screen "Lists" 1440x900, template "Tpl"
   TextField "frm_1" at 12,128 size 1416x70; Text 'Text'
   TextField "txt_1" at 21,132 size 300x23; Text 'POSTAVKE (dok sustav stoji)'
   TextField "txt_2" at 21,162 size 120x28; Text 'Redoslijed'
   SymbolicIOField "sym_1" at 141,162 size 248x28; TextOff '0'; TextOn '1'; TextList "TL_Order"
      ProcessValue <- "CfgOrderMode"
   TextField "txt_3" at 420,162 size 218x28; Text 'SEMI: transfer po koraku'
   SymbolicIOField "sym_2" at 638,162 size 82x28; TextOff '0'; TextOn '1'; TextList "TL_YesNo"
      ProcessValue <- "CfgSemiPerTransfer"
   TextField "txt_4" at 750,162 size 135x28; Text 'Ravnoteža'
   SymbolicIOField "sym_3" at 885,162 size 195x28; TextOff '0'; TextOn '1'; TextList "TL_BalMode"
      ProcessValue <- "CfgBalMode"
   TextField "txt_5" at 1110,162 size 60x28; Text 'Istovar'
   IOField "io_1" at 1170,162 size 45x28; FormatPattern 99
      ProcessValue <- "UTotal"
   TextField "txt_6" at 1230,162 size 60x28; Text 'Ukrcaj'
   IOField "io_2" at 1290,162 size 45x28; FormatPattern 99
      ProcessValue <- "LTotal"
   TextField "txt_7" at 12,210 size 350x23; Text 'LISTA ZA ISTOVAR (DB20) 1-24'
   TextField "txt_8" at 12,238 size 34x22; Text '1'
   IOField "io_3" at 51,238 size 68x22; FormatPattern 999
      ProcessValue <- "UList_01"
   SymbolicIOField "sym_4" at 123,238 size 112x22; TextOff '0'; TextOn '1'; TextList "TL_ListSt"
      ProcessValue <- "UState_01"
   TextField "txt_9" at 12,263 size 34x22; Text '2'
   IOField "io_4" at 51,263 size 68x22; FormatPattern 999
      ProcessValue <- "UList_02"
   SymbolicIOField "sym_5" at 123,263 size 112x22; TextOff '0'; TextOn '1'; TextList "TL_ListSt"
      ProcessValue <- "UState_02"
   TextField "txt_10" at 12,288 size 34x22; Text '3'
   IOField "io_5" at 51,288 size 68x22; FormatPattern 999
      ProcessValue <- "UList_03"
   SymbolicIOField "sym_6" at 123,288 size 112x22; TextOff '0'; TextOn '1'; TextList "TL_ListSt"
      ProcessValue <- "UState_03"
   TextField "txt_11" at 12,313 size 34x22; Text '4'
   IOField "io_6" at 51,313 size 68x22; FormatPattern 999
      ProcessValue <- "UList_04"
   SymbolicIOField "sym_7" at 123,313 size 112x22; TextOff '0'; TextOn '1'; TextList "TL_ListSt"
      ProcessValue <- "UState_04"
   TextField "txt_12" at 12,338 size 34x22; Text '5'
   IOField "io_7" at 51,338 size 68x22; FormatPattern 999
      ProcessValue <- "UList_05"
   SymbolicIOField "sym_8" at 123,338 size 112x22; TextOff '0'; TextOn '1'; TextList "TL_ListSt"
      ProcessValue <- "UState_05"
   TextField "txt_13" at 12,363 size 34x22; Text '6'
   IOField "io_8" at 51,363 size 68x22; FormatPattern 999
      ProcessValue <- "UList_06"
   SymbolicIOField "sym_9" at 123,363 size 112x22; TextOff '0'; TextOn '1'; TextList "TL_ListSt"
      ProcessValue <- "UState_06"
   TextField "txt_14" at 12,388 size 34x22; Text '7'
   IOField "io_9" at 51,388 size 68x22; FormatPattern 999
      ProcessValue <- "UList_07"
   SymbolicIOField "sym_10" at 123,388 size 112x22; TextOff '0'; TextOn '1'; TextList "TL_ListSt"
      ProcessValue <- "UState_07"
   TextField "txt_15" at 12,413 size 34x22; Text '8'
   IOField "io_10" at 51,413 size 68x22; FormatPattern 999
      ProcessValue <- "UList_08"
   SymbolicIOField "sym_11" at 123,413 size 112x22; TextOff '0'; TextOn '1'; TextList "TL_ListSt"
      ProcessValue <- "UState_08"
   TextField "txt_16" at 12,438 size 34x22; Text '9'
   IOField "io_11" at 51,438 size 68x22; FormatPattern 999
      ProcessValue <- "UList_09"
   SymbolicIOField "sym_12" at 123,438 size 112x22; TextOff '0'; TextOn '1'; TextList "TL_ListSt"
      ProcessValue <- "UState_09"
   TextField "txt_17" at 12,463 size 34x22; Text '10'
   IOField "io_12" at 51,463 size 68x22; FormatPattern 999
      ProcessValue <- "UList_10"
   SymbolicIOField "sym_13" at 123,463 size 112x22; TextOff '0'; TextOn '1'; TextList "TL_ListSt"
      ProcessValue <- "UState_10"
   TextField "txt_18" at 12,488 size 34x22; Text '11'
   IOField "io_13" at 51,488 size 68x22; FormatPattern 999
      ProcessValue <- "UList_11"
   SymbolicIOField "sym_14" at 123,488 size 112x22; TextOff '0'; TextOn '1'; TextList "TL_ListSt"
      ProcessValue <- "UState_11"
   TextField "txt_19" at 12,513 size 34x22; Text '12'
   IOField "io_14" at 51,513 size 68x22; FormatPattern 999
      ProcessValue <- "UList_12"
   SymbolicIOField "sym_15" at 123,513 size 112x22; TextOff '0'; TextOn '1'; TextList "TL_ListSt"
      ProcessValue <- "UState_12"
   TextField "txt_20" at 12,538 size 34x22; Text '13'
   IOField "io_15" at 51,538 size 68x22; FormatPattern 999
      ProcessValue <- "UList_13"
   SymbolicIOField "sym_16" at 123,538 size 112x22; TextOff '0'; TextOn '1'; TextList "TL_ListSt"
      ProcessValue <- "UState_13"
   TextField "txt_21" at 12,563 size 34x22; Text '14'
   IOField "io_16" at 51,563 size 68x22; FormatPattern 999
      ProcessValue <- "UList_14"
   SymbolicIOField "sym_17" at 123,563 size 112x22; TextOff '0'; TextOn '1'; TextList "TL_ListSt"
      ProcessValue <- "UState_14"
   TextField "txt_22" at 12,588 size 34x22; Text '15'
   IOField "io_17" at 51,588 size 68x22; FormatPattern 999
      ProcessValue <- "UList_15"
   SymbolicIOField "sym_18" at 123,588 size 112x22; TextOff '0'; TextOn '1'; TextList "TL_ListSt"
      ProcessValue <- "UState_15"
   TextField "txt_23" at 12,613 size 34x22; Text '16'
   IOField "io_18" at 51,613 size 68x22; FormatPattern 999
      ProcessValue <- "UList_16"
   SymbolicIOField "sym_19" at 123,613 size 112x22; TextOff '0'; TextOn '1'; TextList "TL_ListSt"
      ProcessValue <- "UState_16"
   TextField "txt_24" at 12,638 size 34x22; Text '17'
   IOField "io_19" at 51,638 size 68x22; FormatPattern 999
      ProcessValue <- "UList_17"
   SymbolicIOField "sym_20" at 123,638 size 112x22; TextOff '0'; TextOn '1'; TextList "TL_ListSt"
      ProcessValue <- "UState_17"
   TextField "txt_25" at 12,663 size 34x22; Text '18'
   IOField "io_20" at 51,663 size 68x22; FormatPattern 999
      ProcessValue <- "UList_18"
   SymbolicIOField "sym_21" at 123,663 size 112x22; TextOff '0'; TextOn '1'; TextList "TL_ListSt"
      ProcessValue <- "UState_18"
   TextField "txt_26" at 12,688 size 34x22; Text '19'
   IOField "io_21" at 51,688 size 68x22; FormatPattern 999
      ProcessValue <- "UList_19"
   SymbolicIOField "sym_22" at 123,688 size 112x22; TextOff '0'; TextOn '1'; TextList "TL_ListSt"
      ProcessValue <- "UState_19"
   TextField "txt_27" at 12,713 size 34x22; Text '20'
   IOField "io_22" at 51,713 size 68x22; FormatPattern 999
      ProcessValue <- "UList_20"
   SymbolicIOField "sym_23" at 123,713 size 112x22; TextOff '0'; TextOn '1'; TextList "TL_ListSt"
      ProcessValue <- "UState_20"
   TextField "txt_28" at 12,738 size 34x22; Text '21'
   IOField "io_23" at 51,738 size 68x22; FormatPattern 999
      ProcessValue <- "UList_21"
   SymbolicIOField "sym_24" at 123,738 size 112x22; TextOff '0'; TextOn '1'; TextList "TL_ListSt"
      ProcessValue <- "UState_21"
   TextField "txt_29" at 12,763 size 34x22; Text '22'
   IOField "io_24" at 51,763 size 68x22; FormatPattern 999
      ProcessValue <- "UList_22"
   SymbolicIOField "sym_25" at 123,763 size 112x22; TextOff '0'; TextOn '1'; TextList "TL_ListSt"
      ProcessValue <- "UState_22"
   TextField "txt_30" at 12,788 size 34x22; Text '23'
   IOField "io_25" at 51,788 size 68x22; FormatPattern 999
      ProcessValue <- "UList_23"
   SymbolicIOField "sym_26" at 123,788 size 112x22; TextOff '0'; TextOn '1'; TextList "TL_ListSt"
      ProcessValue <- "UState_23"
   TextField "txt_31" at 12,813 size 34x22; Text '24'
   IOField "io_26" at 51,813 size 68x22; FormatPattern 999
      ProcessValue <- "UList_24"
   SymbolicIOField "sym_27" at 123,813 size 112x22; TextOff '0'; TextOn '1'; TextList "TL_ListSt"
      ProcessValue <- "UState_24"
   TextField "txt_32" at 368,210 size 350x23; Text 'LISTA ZA ISTOVAR 25-48'
   TextField "txt_33" at 368,238 size 34x22; Text '25'
   IOField "io_27" at 406,238 size 68x22; FormatPattern 999
      ProcessValue <- "UList_25"
   SymbolicIOField "sym_28" at 478,238 size 112x22; TextOff '0'; TextOn '1'; TextList "TL_ListSt"
      ProcessValue <- "UState_25"
   TextField "txt_34" at 368,263 size 34x22; Text '26'
   IOField "io_28" at 406,263 size 68x22; FormatPattern 999
      ProcessValue <- "UList_26"
   SymbolicIOField "sym_29" at 478,263 size 112x22; TextOff '0'; TextOn '1'; TextList "TL_ListSt"
      ProcessValue <- "UState_26"
   TextField "txt_35" at 368,288 size 34x22; Text '27'
   IOField "io_29" at 406,288 size 68x22; FormatPattern 999
      ProcessValue <- "UList_27"
   SymbolicIOField "sym_30" at 478,288 size 112x22; TextOff '0'; TextOn '1'; TextList "TL_ListSt"
      ProcessValue <- "UState_27"
   TextField "txt_36" at 368,313 size 34x22; Text '28'
   IOField "io_30" at 406,313 size 68x22; FormatPattern 999
      ProcessValue <- "UList_28"
   SymbolicIOField "sym_31" at 478,313 size 112x22; TextOff '0'; TextOn '1'; TextList "TL_ListSt"
      ProcessValue <- "UState_28"
   TextField "txt_37" at 368,338 size 34x22; Text '29'
   IOField "io_31" at 406,338 size 68x22; FormatPattern 999
      ProcessValue <- "UList_29"
   SymbolicIOField "sym_32" at 478,338 size 112x22; TextOff '0'; TextOn '1'; TextList "TL_ListSt"
      ProcessValue <- "UState_29"
   TextField "txt_38" at 368,363 size 34x22; Text '30'
   IOField "io_32" at 406,363 size 68x22; FormatPattern 999
      ProcessValue <- "UList_30"
   SymbolicIOField "sym_33" at 478,363 size 112x22; TextOff '0'; TextOn '1'; TextList "TL_ListSt"
      ProcessValue <- "UState_30"
   TextField "txt_39" at 368,388 size 34x22; Text '31'
   IOField "io_33" at 406,388 size 68x22; FormatPattern 999
      ProcessValue <- "UList_31"
   SymbolicIOField "sym_34" at 478,388 size 112x22; TextOff '0'; TextOn '1'; TextList "TL_ListSt"
      ProcessValue <- "UState_31"
   TextField "txt_40" at 368,413 size 34x22; Text '32'
   IOField "io_34" at 406,413 size 68x22; FormatPattern 999
      ProcessValue <- "UList_32"
   SymbolicIOField "sym_35" at 478,413 size 112x22; TextOff '0'; TextOn '1'; TextList "TL_ListSt"
      ProcessValue <- "UState_32"
   TextField "txt_41" at 368,438 size 34x22; Text '33'
   IOField "io_35" at 406,438 size 68x22; FormatPattern 999
      ProcessValue <- "UList_33"
   SymbolicIOField "sym_36" at 478,438 size 112x22; TextOff '0'; TextOn '1'; TextList "TL_ListSt"
      ProcessValue <- "UState_33"
   TextField "txt_42" at 368,463 size 34x22; Text '34'
   IOField "io_36" at 406,463 size 68x22; FormatPattern 999
      ProcessValue <- "UList_34"
   SymbolicIOField "sym_37" at 478,463 size 112x22; TextOff '0'; TextOn '1'; TextList "TL_ListSt"
      ProcessValue <- "UState_34"
   TextField "txt_43" at 368,488 size 34x22; Text '35'
   IOField "io_37" at 406,488 size 68x22; FormatPattern 999
      ProcessValue <- "UList_35"
   SymbolicIOField "sym_38" at 478,488 size 112x22; TextOff '0'; TextOn '1'; TextList "TL_ListSt"
      ProcessValue <- "UState_35"
   TextField "txt_44" at 368,513 size 34x22; Text '36'
   IOField "io_38" at 406,513 size 68x22; FormatPattern 999
      ProcessValue <- "UList_36"
   SymbolicIOField "sym_39" at 478,513 size 112x22; TextOff '0'; TextOn '1'; TextList "TL_ListSt"
      ProcessValue <- "UState_36"
   TextField "txt_45" at 368,538 size 34x22; Text '37'
   IOField "io_39" at 406,538 size 68x22; FormatPattern 999
      ProcessValue <- "UList_37"
   SymbolicIOField "sym_40" at 478,538 size 112x22; TextOff '0'; TextOn '1'; TextList "TL_ListSt"
      ProcessValue <- "UState_37"
   TextField "txt_46" at 368,563 size 34x22; Text '38'
   IOField "io_40" at 406,563 size 68x22; FormatPattern 999
      ProcessValue <- "UList_38"
   SymbolicIOField "sym_41" at 478,563 size 112x22; TextOff '0'; TextOn '1'; TextList "TL_ListSt"
      ProcessValue <- "UState_38"
   TextField "txt_47" at 368,588 size 34x22; Text '39'
   IOField "io_41" at 406,588 size 68x22; FormatPattern 999
      ProcessValue <- "UList_39"
   SymbolicIOField "sym_42" at 478,588 size 112x22; TextOff '0'; TextOn '1'; TextList "TL_ListSt"
      ProcessValue <- "UState_39"
   TextField "txt_48" at 368,613 size 34x22; Text '40'
   IOField "io_42" at 406,613 size 68x22; FormatPattern 999
      ProcessValue <- "UList_40"
   SymbolicIOField "sym_43" at 478,613 size 112x22; TextOff '0'; TextOn '1'; TextList "TL_ListSt"
      ProcessValue <- "UState_40"
   TextField "txt_49" at 368,638 size 34x22; Text '41'
   IOField "io_43" at 406,638 size 68x22; FormatPattern 999
      ProcessValue <- "UList_41"
   SymbolicIOField "sym_44" at 478,638 size 112x22; TextOff '0'; TextOn '1'; TextList "TL_ListSt"
      ProcessValue <- "UState_41"
   TextField "txt_50" at 368,663 size 34x22; Text '42'
   IOField "io_44" at 406,663 size 68x22; FormatPattern 999
      ProcessValue <- "UList_42"
   SymbolicIOField "sym_45" at 478,663 size 112x22; TextOff '0'; TextOn '1'; TextList "TL_ListSt"
      ProcessValue <- "UState_42"
   TextField "txt_51" at 368,688 size 34x22; Text '43'
   IOField "io_45" at 406,688 size 68x22; FormatPattern 999
      ProcessValue <- "UList_43"
   SymbolicIOField "sym_46" at 478,688 size 112x22; TextOff '0'; TextOn '1'; TextList "TL_ListSt"
      ProcessValue <- "UState_43"
   TextField "txt_52" at 368,713 size 34x22; Text '44'
   IOField "io_46" at 406,713 size 68x22; FormatPattern 999
      ProcessValue <- "UList_44"
   SymbolicIOField "sym_47" at 478,713 size 112x22; TextOff '0'; TextOn '1'; TextList "TL_ListSt"
      ProcessValue <- "UState_44"
   TextField "txt_53" at 368,738 size 34x22; Text '45'
   IOField "io_47" at 406,738 size 68x22; FormatPattern 999
      ProcessValue <- "UList_45"
   SymbolicIOField "sym_48" at 478,738 size 112x22; TextOff '0'; TextOn '1'; TextList "TL_ListSt"
      ProcessValue <- "UState_45"
   TextField "txt_54" at 368,763 size 34x22; Text '46'
   IOField "io_48" at 406,763 size 68x22; FormatPattern 999
      ProcessValue <- "UList_46"
   SymbolicIOField "sym_49" at 478,763 size 112x22; TextOff '0'; TextOn '1'; TextList "TL_ListSt"
      ProcessValue <- "UState_46"
   TextField "txt_55" at 368,788 size 34x22; Text '47'
   IOField "io_49" at 406,788 size 68x22; FormatPattern 999
      ProcessValue <- "UList_47"
   SymbolicIOField "sym_50" at 478,788 size 112x22; TextOff '0'; TextOn '1'; TextList "TL_ListSt"
      ProcessValue <- "UState_47"
   TextField "txt_56" at 368,813 size 34x22; Text '48'
   IOField "io_50" at 406,813 size 68x22; FormatPattern 999
      ProcessValue <- "UList_48"
   SymbolicIOField "sym_51" at 478,813 size 112x22; TextOff '0'; TextOn '1'; TextList "TL_ListSt"
      ProcessValue <- "UState_48"
   TextField "txt_57" at 723,210 size 350x23; Text 'LISTA ZA UKRCAJ (DB21) 1-24'
   TextField "txt_58" at 723,238 size 34x22; Text '1'
   IOField "io_51" at 762,238 size 68x22; FormatPattern 999
      ProcessValue <- "LList_01"
   SymbolicIOField "sym_52" at 834,238 size 112x22; TextOff '0'; TextOn '1'; TextList "TL_ListSt"
      ProcessValue <- "LState_01"
   TextField "txt_59" at 723,263 size 34x22; Text '2'
   IOField "io_52" at 762,263 size 68x22; FormatPattern 999
      ProcessValue <- "LList_02"
   SymbolicIOField "sym_53" at 834,263 size 112x22; TextOff '0'; TextOn '1'; TextList "TL_ListSt"
      ProcessValue <- "LState_02"
   TextField "txt_60" at 723,288 size 34x22; Text '3'
   IOField "io_53" at 762,288 size 68x22; FormatPattern 999
      ProcessValue <- "LList_03"
   SymbolicIOField "sym_54" at 834,288 size 112x22; TextOff '0'; TextOn '1'; TextList "TL_ListSt"
      ProcessValue <- "LState_03"
   TextField "txt_61" at 723,313 size 34x22; Text '4'
   IOField "io_54" at 762,313 size 68x22; FormatPattern 999
      ProcessValue <- "LList_04"
   SymbolicIOField "sym_55" at 834,313 size 112x22; TextOff '0'; TextOn '1'; TextList "TL_ListSt"
      ProcessValue <- "LState_04"
   TextField "txt_62" at 723,338 size 34x22; Text '5'
   IOField "io_55" at 762,338 size 68x22; FormatPattern 999
      ProcessValue <- "LList_05"
   SymbolicIOField "sym_56" at 834,338 size 112x22; TextOff '0'; TextOn '1'; TextList "TL_ListSt"
      ProcessValue <- "LState_05"
   TextField "txt_63" at 723,363 size 34x22; Text '6'
   IOField "io_56" at 762,363 size 68x22; FormatPattern 999
      ProcessValue <- "LList_06"
   SymbolicIOField "sym_57" at 834,363 size 112x22; TextOff '0'; TextOn '1'; TextList "TL_ListSt"
      ProcessValue <- "LState_06"
   TextField "txt_64" at 723,388 size 34x22; Text '7'
   IOField "io_57" at 762,388 size 68x22; FormatPattern 999
      ProcessValue <- "LList_07"
   SymbolicIOField "sym_58" at 834,388 size 112x22; TextOff '0'; TextOn '1'; TextList "TL_ListSt"
      ProcessValue <- "LState_07"
   TextField "txt_65" at 723,413 size 34x22; Text '8'
   IOField "io_58" at 762,413 size 68x22; FormatPattern 999
      ProcessValue <- "LList_08"
   SymbolicIOField "sym_59" at 834,413 size 112x22; TextOff '0'; TextOn '1'; TextList "TL_ListSt"
      ProcessValue <- "LState_08"
   TextField "txt_66" at 723,438 size 34x22; Text '9'
   IOField "io_59" at 762,438 size 68x22; FormatPattern 999
      ProcessValue <- "LList_09"
   SymbolicIOField "sym_60" at 834,438 size 112x22; TextOff '0'; TextOn '1'; TextList "TL_ListSt"
      ProcessValue <- "LState_09"
   TextField "txt_67" at 723,463 size 34x22; Text '10'
   IOField "io_60" at 762,463 size 68x22; FormatPattern 999
      ProcessValue <- "LList_10"
   SymbolicIOField "sym_61" at 834,463 size 112x22; TextOff '0'; TextOn '1'; TextList "TL_ListSt"
      ProcessValue <- "LState_10"
   TextField "txt_68" at 723,488 size 34x22; Text '11'
   IOField "io_61" at 762,488 size 68x22; FormatPattern 999
      ProcessValue <- "LList_11"
   SymbolicIOField "sym_62" at 834,488 size 112x22; TextOff '0'; TextOn '1'; TextList "TL_ListSt"
      ProcessValue <- "LState_11"
   TextField "txt_69" at 723,513 size 34x22; Text '12'
   IOField "io_62" at 762,513 size 68x22; FormatPattern 999
      ProcessValue <- "LList_12"
   SymbolicIOField "sym_63" at 834,513 size 112x22; TextOff '0'; TextOn '1'; TextList "TL_ListSt"
      ProcessValue <- "LState_12"
   TextField "txt_70" at 723,538 size 34x22; Text '13'
   IOField "io_63" at 762,538 size 68x22; FormatPattern 999
      ProcessValue <- "LList_13"
   SymbolicIOField "sym_64" at 834,538 size 112x22; TextOff '0'; TextOn '1'; TextList "TL_ListSt"
      ProcessValue <- "LState_13"
   TextField "txt_71" at 723,563 size 34x22; Text '14'
   IOField "io_64" at 762,563 size 68x22; FormatPattern 999
      ProcessValue <- "LList_14"
   SymbolicIOField "sym_65" at 834,563 size 112x22; TextOff '0'; TextOn '1'; TextList "TL_ListSt"
      ProcessValue <- "LState_14"
   TextField "txt_72" at 723,588 size 34x22; Text '15'
   IOField "io_65" at 762,588 size 68x22; FormatPattern 999
      ProcessValue <- "LList_15"
   SymbolicIOField "sym_66" at 834,588 size 112x22; TextOff '0'; TextOn '1'; TextList "TL_ListSt"
      ProcessValue <- "LState_15"
   TextField "txt_73" at 723,613 size 34x22; Text '16'
   IOField "io_66" at 762,613 size 68x22; FormatPattern 999
      ProcessValue <- "LList_16"
   SymbolicIOField "sym_67" at 834,613 size 112x22; TextOff '0'; TextOn '1'; TextList "TL_ListSt"
      ProcessValue <- "LState_16"
   TextField "txt_74" at 723,638 size 34x22; Text '17'
   IOField "io_67" at 762,638 size 68x22; FormatPattern 999
      ProcessValue <- "LList_17"
   SymbolicIOField "sym_68" at 834,638 size 112x22; TextOff '0'; TextOn '1'; TextList "TL_ListSt"
      ProcessValue <- "LState_17"
   TextField "txt_75" at 723,663 size 34x22; Text '18'
   IOField "io_68" at 762,663 size 68x22; FormatPattern 999
      ProcessValue <- "LList_18"
   SymbolicIOField "sym_69" at 834,663 size 112x22; TextOff '0'; TextOn '1'; TextList "TL_ListSt"
      ProcessValue <- "LState_18"
   TextField "txt_76" at 723,688 size 34x22; Text '19'
   IOField "io_69" at 762,688 size 68x22; FormatPattern 999
      ProcessValue <- "LList_19"
   SymbolicIOField "sym_70" at 834,688 size 112x22; TextOff '0'; TextOn '1'; TextList "TL_ListSt"
      ProcessValue <- "LState_19"
   TextField "txt_77" at 723,713 size 34x22; Text '20'
   IOField "io_70" at 762,713 size 68x22; FormatPattern 999
      ProcessValue <- "LList_20"
   SymbolicIOField "sym_71" at 834,713 size 112x22; TextOff '0'; TextOn '1'; TextList "TL_ListSt"
      ProcessValue <- "LState_20"
   TextField "txt_78" at 723,738 size 34x22; Text '21'
   IOField "io_71" at 762,738 size 68x22; FormatPattern 999
      ProcessValue <- "LList_21"
   SymbolicIOField "sym_72" at 834,738 size 112x22; TextOff '0'; TextOn '1'; TextList "TL_ListSt"
      ProcessValue <- "LState_21"
   TextField "txt_79" at 723,763 size 34x22; Text '22'
   IOField "io_72" at 762,763 size 68x22; FormatPattern 999
      ProcessValue <- "LList_22"
   SymbolicIOField "sym_73" at 834,763 size 112x22; TextOff '0'; TextOn '1'; TextList "TL_ListSt"
      ProcessValue <- "LState_22"
   TextField "txt_80" at 723,788 size 34x22; Text '23'
   IOField "io_73" at 762,788 size 68x22; FormatPattern 999
      ProcessValue <- "LList_23"
   SymbolicIOField "sym_74" at 834,788 size 112x22; TextOff '0'; TextOn '1'; TextList "TL_ListSt"
      ProcessValue <- "LState_23"
   TextField "txt_81" at 723,813 size 34x22; Text '24'
   IOField "io_74" at 762,813 size 68x22; FormatPattern 999
      ProcessValue <- "LList_24"
   SymbolicIOField "sym_75" at 834,813 size 112x22; TextOff '0'; TextOn '1'; TextList "TL_ListSt"
      ProcessValue <- "LState_24"
   TextField "txt_82" at 1078,210 size 350x23; Text 'LISTA ZA UKRCAJ 25-48'
   TextField "txt_83" at 1078,238 size 34x22; Text '25'
   IOField "io_75" at 1118,238 size 68x22; FormatPattern 999
      ProcessValue <- "LList_25"
   SymbolicIOField "sym_76" at 1190,238 size 112x22; TextOff '0'; TextOn '1'; TextList "TL_ListSt"
      ProcessValue <- "LState_25"
   TextField "txt_84" at 1078,263 size 34x22; Text '26'
   IOField "io_76" at 1118,263 size 68x22; FormatPattern 999
      ProcessValue <- "LList_26"
   SymbolicIOField "sym_77" at 1190,263 size 112x22; TextOff '0'; TextOn '1'; TextList "TL_ListSt"
      ProcessValue <- "LState_26"
   TextField "txt_85" at 1078,288 size 34x22; Text '27'
   IOField "io_77" at 1118,288 size 68x22; FormatPattern 999
      ProcessValue <- "LList_27"
   SymbolicIOField "sym_78" at 1190,288 size 112x22; TextOff '0'; TextOn '1'; TextList "TL_ListSt"
      ProcessValue <- "LState_27"
   TextField "txt_86" at 1078,313 size 34x22; Text '28'
   IOField "io_78" at 1118,313 size 68x22; FormatPattern 999
      ProcessValue <- "LList_28"
   SymbolicIOField "sym_79" at 1190,313 size 112x22; TextOff '0'; TextOn '1'; TextList "TL_ListSt"
      ProcessValue <- "LState_28"
   TextField "txt_87" at 1078,338 size 34x22; Text '29'
   IOField "io_79" at 1118,338 size 68x22; FormatPattern 999
      ProcessValue <- "LList_29"
   SymbolicIOField "sym_80" at 1190,338 size 112x22; TextOff '0'; TextOn '1'; TextList "TL_ListSt"
      ProcessValue <- "LState_29"
   TextField "txt_88" at 1078,363 size 34x22; Text '30'
   IOField "io_80" at 1118,363 size 68x22; FormatPattern 999
      ProcessValue <- "LList_30"
   SymbolicIOField "sym_81" at 1190,363 size 112x22; TextOff '0'; TextOn '1'; TextList "TL_ListSt"
      ProcessValue <- "LState_30"
   TextField "txt_89" at 1078,388 size 34x22; Text '31'
   IOField "io_81" at 1118,388 size 68x22; FormatPattern 999
      ProcessValue <- "LList_31"
   SymbolicIOField "sym_82" at 1190,388 size 112x22; TextOff '0'; TextOn '1'; TextList "TL_ListSt"
      ProcessValue <- "LState_31"
   TextField "txt_90" at 1078,413 size 34x22; Text '32'
   IOField "io_82" at 1118,413 size 68x22; FormatPattern 999
      ProcessValue <- "LList_32"
   SymbolicIOField "sym_83" at 1190,413 size 112x22; TextOff '0'; TextOn '1'; TextList "TL_ListSt"
      ProcessValue <- "LState_32"
   TextField "txt_91" at 1078,438 size 34x22; Text '33'
   IOField "io_83" at 1118,438 size 68x22; FormatPattern 999
      ProcessValue <- "LList_33"
   SymbolicIOField "sym_84" at 1190,438 size 112x22; TextOff '0'; TextOn '1'; TextList "TL_ListSt"
      ProcessValue <- "LState_33"
   TextField "txt_92" at 1078,463 size 34x22; Text '34'
   IOField "io_84" at 1118,463 size 68x22; FormatPattern 999
      ProcessValue <- "LList_34"
   SymbolicIOField "sym_85" at 1190,463 size 112x22; TextOff '0'; TextOn '1'; TextList "TL_ListSt"
      ProcessValue <- "LState_34"
   TextField "txt_93" at 1078,488 size 34x22; Text '35'
   IOField "io_85" at 1118,488 size 68x22; FormatPattern 999
      ProcessValue <- "LList_35"
   SymbolicIOField "sym_86" at 1190,488 size 112x22; TextOff '0'; TextOn '1'; TextList "TL_ListSt"
      ProcessValue <- "LState_35"
   TextField "txt_94" at 1078,513 size 34x22; Text '36'
   IOField "io_86" at 1118,513 size 68x22; FormatPattern 999
      ProcessValue <- "LList_36"
   SymbolicIOField "sym_87" at 1190,513 size 112x22; TextOff '0'; TextOn '1'; TextList "TL_ListSt"
      ProcessValue <- "LState_36"
   TextField "txt_95" at 1078,538 size 34x22; Text '37'
   IOField "io_87" at 1118,538 size 68x22; FormatPattern 999
      ProcessValue <- "LList_37"
   SymbolicIOField "sym_88" at 1190,538 size 112x22; TextOff '0'; TextOn '1'; TextList "TL_ListSt"
      ProcessValue <- "LState_37"
   TextField "txt_96" at 1078,563 size 34x22; Text '38'
   IOField "io_88" at 1118,563 size 68x22; FormatPattern 999
      ProcessValue <- "LList_38"
   SymbolicIOField "sym_89" at 1190,563 size 112x22; TextOff '0'; TextOn '1'; TextList "TL_ListSt"
      ProcessValue <- "LState_38"
   TextField "txt_97" at 1078,588 size 34x22; Text '39'
   IOField "io_89" at 1118,588 size 68x22; FormatPattern 999
      ProcessValue <- "LList_39"
   SymbolicIOField "sym_90" at 1190,588 size 112x22; TextOff '0'; TextOn '1'; TextList "TL_ListSt"
      ProcessValue <- "LState_39"
   TextField "txt_98" at 1078,613 size 34x22; Text '40'
   IOField "io_90" at 1118,613 size 68x22; FormatPattern 999
      ProcessValue <- "LList_40"
   SymbolicIOField "sym_91" at 1190,613 size 112x22; TextOff '0'; TextOn '1'; TextList "TL_ListSt"
      ProcessValue <- "LState_40"
   TextField "txt_99" at 1078,638 size 34x22; Text '41'
   IOField "io_91" at 1118,638 size 68x22; FormatPattern 999
      ProcessValue <- "LList_41"
   SymbolicIOField "sym_92" at 1190,638 size 112x22; TextOff '0'; TextOn '1'; TextList "TL_ListSt"
      ProcessValue <- "LState_41"
   TextField "txt_100" at 1078,663 size 34x22; Text '42'
   IOField "io_92" at 1118,663 size 68x22; FormatPattern 999
      ProcessValue <- "LList_42"
   SymbolicIOField "sym_93" at 1190,663 size 112x22; TextOff '0'; TextOn '1'; TextList "TL_ListSt"
      ProcessValue <- "LState_42"
   TextField "txt_101" at 1078,688 size 34x22; Text '43'
   IOField "io_93" at 1118,688 size 68x22; FormatPattern 999
      ProcessValue <- "LList_43"
   SymbolicIOField "sym_94" at 1190,688 size 112x22; TextOff '0'; TextOn '1'; TextList "TL_ListSt"
      ProcessValue <- "LState_43"
   TextField "txt_102" at 1078,713 size 34x22; Text '44'
   IOField "io_94" at 1118,713 size 68x22; FormatPattern 999
      ProcessValue <- "LList_44"
   SymbolicIOField "sym_95" at 1190,713 size 112x22; TextOff '0'; TextOn '1'; TextList "TL_ListSt"
      ProcessValue <- "LState_44"
   TextField "txt_103" at 1078,738 size 34x22; Text '45'
   IOField "io_95" at 1118,738 size 68x22; FormatPattern 999
      ProcessValue <- "LList_45"
   SymbolicIOField "sym_96" at 1190,738 size 112x22; TextOff '0'; TextOn '1'; TextList "TL_ListSt"
      ProcessValue <- "LState_45"
   TextField "txt_104" at 1078,763 size 34x22; Text '46'
   IOField "io_96" at 1118,763 size 68x22; FormatPattern 999
      ProcessValue <- "LList_46"
   SymbolicIOField "sym_97" at 1190,763 size 112x22; TextOff '0'; TextOn '1'; TextList "TL_ListSt"
      ProcessValue <- "LState_46"
   TextField "txt_105" at 1078,788 size 34x22; Text '47'
   IOField "io_97" at 1118,788 size 68x22; FormatPattern 999
      ProcessValue <- "LList_47"
   SymbolicIOField "sym_98" at 1190,788 size 112x22; TextOff '0'; TextOn '1'; TextList "TL_ListSt"
      ProcessValue <- "LState_47"
   TextField "txt_106" at 1078,813 size 34x22; Text '48'
   IOField "io_98" at 1118,813 size 68x22; FormatPattern 999
      ProcessValue <- "LList_48"
   SymbolicIOField "sym_99" at 1190,813 size 112x22; TextOff '0'; TextOn '1'; TextList "TL_ListSt"
      ProcessValue <- "LState_48"

screen "Manual" 1440x900, template "Tpl"
   TextField "txt_1" at 45,128 size 334x23; Text 'BAY 1 - SKLADIŠTE (yard)'
   TextField "txt_2" at 558,128 size 334x23; Text 'BAY 0 - BROD (ship)'
   TextField "frm_1" at 42,155 size 854x30; Text 'Text'
   TextField "frm_2" at 417,187 size 105x602; Text 'Text'
   TextField "txt_3" at 417,792 size 105x18; Text 'OBALA / kran y'
   TextField "frm_3" at 39,183 size 346x608; Text 'Text'
   TextField "frm_4" at 552,183 size 346x608; Text 'Text'
   TextField "frm_5" at 724,183 size 3x608; Text 'Text'
   TextField "txt_4" at 12,203 size 30x18; Text 'y0'
   TextField "txt_5" at 12,253 size 30x18; Text 'y1'
   TextField "txt_6" at 12,303 size 30x18; Text 'y2'
   TextField "txt_7" at 12,353 size 30x18; Text 'y3'
   TextField "txt_8" at 12,403 size 30x18; Text 'y4'
   TextField "txt_9" at 12,453 size 30x18; Text 'y5'
   TextField "txt_10" at 12,503 size 30x18; Text 'y6'
   TextField "txt_11" at 12,553 size 30x18; Text 'y7'
   TextField "txt_12" at 12,603 size 30x18; Text 'y8'
   TextField "txt_13" at 12,653 size 30x18; Text 'y9'
   TextField "txt_14" at 12,703 size 30x18; Text 'y10'
   TextField "txt_15" at 12,753 size 30x18; Text 'y11'
   TextField "txt_16" at 45,793 size 78x17; Text 'x0'
   TextField "txt_17" at 130,793 size 78x17; Text 'x1'
   TextField "txt_18" at 216,793 size 78x17; Text 'x2'
   TextField "txt_19" at 302,793 size 78x17; Text 'x3'
   TextField "txt_20" at 558,793 size 78x17; Text 'x0'
   TextField "txt_21" at 644,793 size 78x17; Text 'x1'
   TextField "txt_22" at 729,793 size 78x17; Text 'x2'
   TextField "txt_23" at 814,793 size 78x17; Text 'x3'
   TextField "txt_24" at 558,813 size 90x23; Text 'LIJEVO'
   IOField "io_1" at 648,813 size 45x23; FormatPattern 99
      ProcessValue <- "BalL"
   TextField "txt_25" at 729,813 size 90x23; Text 'DESNO'
   IOField "io_2" at 819,813 size 45x23; FormatPattern 99
      ProcessValue <- "BalR"
   Rectangle "cel_1" at 45,190 size 78x45
      Appearance <- "CellSt1_00"
   IOField "io_3" at 50,196 size 68x33; FormatPattern 999
      ProcessValue <- "Cell1_00"
      Appearance <- "CellSt1_00"
   Rectangle "cel_2" at 45,240 size 78x45
      Appearance <- "CellSt1_01"
   IOField "io_4" at 50,246 size 68x33; FormatPattern 999
      ProcessValue <- "Cell1_01"
      Appearance <- "CellSt1_01"
   Rectangle "cel_3" at 45,290 size 78x45
      Appearance <- "CellSt1_02"
   IOField "io_5" at 50,296 size 68x33; FormatPattern 999
      ProcessValue <- "Cell1_02"
      Appearance <- "CellSt1_02"
   Rectangle "cel_4" at 45,340 size 78x45
      Appearance <- "CellSt1_03"
   IOField "io_6" at 50,346 size 68x33; FormatPattern 999
      ProcessValue <- "Cell1_03"
      Appearance <- "CellSt1_03"
   Rectangle "cel_5" at 45,390 size 78x45
      Appearance <- "CellSt1_04"
   IOField "io_7" at 50,396 size 68x33; FormatPattern 999
      ProcessValue <- "Cell1_04"
      Appearance <- "CellSt1_04"
   Rectangle "cel_6" at 45,440 size 78x45
      Appearance <- "CellSt1_05"
   IOField "io_8" at 50,446 size 68x33; FormatPattern 999
      ProcessValue <- "Cell1_05"
      Appearance <- "CellSt1_05"
   Rectangle "cel_7" at 45,490 size 78x45
      Appearance <- "CellSt1_06"
   IOField "io_9" at 50,496 size 68x33; FormatPattern 999
      ProcessValue <- "Cell1_06"
      Appearance <- "CellSt1_06"
   Rectangle "cel_8" at 45,540 size 78x45
      Appearance <- "CellSt1_07"
   IOField "io_10" at 50,546 size 68x33; FormatPattern 999
      ProcessValue <- "Cell1_07"
      Appearance <- "CellSt1_07"
   Rectangle "cel_9" at 45,590 size 78x45
      Appearance <- "CellSt1_08"
   IOField "io_11" at 50,596 size 68x33; FormatPattern 999
      ProcessValue <- "Cell1_08"
      Appearance <- "CellSt1_08"
   Rectangle "cel_10" at 45,640 size 78x45
      Appearance <- "CellSt1_09"
   IOField "io_12" at 50,646 size 68x33; FormatPattern 999
      ProcessValue <- "Cell1_09"
      Appearance <- "CellSt1_09"
   Rectangle "cel_11" at 45,690 size 78x45
      Appearance <- "CellSt1_10"
   IOField "io_13" at 50,696 size 68x33; FormatPattern 999
      ProcessValue <- "Cell1_10"
      Appearance <- "CellSt1_10"
   Rectangle "cel_12" at 45,740 size 78x45
      Appearance <- "CellSt1_11"
   IOField "io_14" at 50,746 size 68x33; FormatPattern 999
      ProcessValue <- "Cell1_11"
      Appearance <- "CellSt1_11"
   Rectangle "cel_13" at 130,190 size 78x45
      Appearance <- "CellSt1_12"
   IOField "io_15" at 136,196 size 68x33; FormatPattern 999
      ProcessValue <- "Cell1_12"
      Appearance <- "CellSt1_12"
   Rectangle "cel_14" at 130,240 size 78x45
      Appearance <- "CellSt1_13"
   IOField "io_16" at 136,246 size 68x33; FormatPattern 999
      ProcessValue <- "Cell1_13"
      Appearance <- "CellSt1_13"
   Rectangle "cel_15" at 130,290 size 78x45
      Appearance <- "CellSt1_14"
   IOField "io_17" at 136,296 size 68x33; FormatPattern 999
      ProcessValue <- "Cell1_14"
      Appearance <- "CellSt1_14"
   Rectangle "cel_16" at 130,340 size 78x45
      Appearance <- "CellSt1_15"
   IOField "io_18" at 136,346 size 68x33; FormatPattern 999
      ProcessValue <- "Cell1_15"
      Appearance <- "CellSt1_15"
   Rectangle "cel_17" at 130,390 size 78x45
      Appearance <- "CellSt1_16"
   IOField "io_19" at 136,396 size 68x33; FormatPattern 999
      ProcessValue <- "Cell1_16"
      Appearance <- "CellSt1_16"
   Rectangle "cel_18" at 130,440 size 78x45
      Appearance <- "CellSt1_17"
   IOField "io_20" at 136,446 size 68x33; FormatPattern 999
      ProcessValue <- "Cell1_17"
      Appearance <- "CellSt1_17"
   Rectangle "cel_19" at 130,490 size 78x45
      Appearance <- "CellSt1_18"
   IOField "io_21" at 136,496 size 68x33; FormatPattern 999
      ProcessValue <- "Cell1_18"
      Appearance <- "CellSt1_18"
   Rectangle "cel_20" at 130,540 size 78x45
      Appearance <- "CellSt1_19"
   IOField "io_22" at 136,546 size 68x33; FormatPattern 999
      ProcessValue <- "Cell1_19"
      Appearance <- "CellSt1_19"
   Rectangle "cel_21" at 130,590 size 78x45
      Appearance <- "CellSt1_20"
   IOField "io_23" at 136,596 size 68x33; FormatPattern 999
      ProcessValue <- "Cell1_20"
      Appearance <- "CellSt1_20"
   Rectangle "cel_22" at 130,640 size 78x45
      Appearance <- "CellSt1_21"
   IOField "io_24" at 136,646 size 68x33; FormatPattern 999
      ProcessValue <- "Cell1_21"
      Appearance <- "CellSt1_21"
   Rectangle "cel_23" at 130,690 size 78x45
      Appearance <- "CellSt1_22"
   IOField "io_25" at 136,696 size 68x33; FormatPattern 999
      ProcessValue <- "Cell1_22"
      Appearance <- "CellSt1_22"
   Rectangle "cel_24" at 130,740 size 78x45
      Appearance <- "CellSt1_23"
   IOField "io_26" at 136,746 size 68x33; FormatPattern 999
      ProcessValue <- "Cell1_23"
      Appearance <- "CellSt1_23"
   Rectangle "cel_25" at 216,190 size 78x45
      Appearance <- "CellSt1_24"
   IOField "io_27" at 221,196 size 68x33; FormatPattern 999
      ProcessValue <- "Cell1_24"
      Appearance <- "CellSt1_24"
   Rectangle "cel_26" at 216,240 size 78x45
      Appearance <- "CellSt1_25"
   IOField "io_28" at 221,246 size 68x33; FormatPattern 999
      ProcessValue <- "Cell1_25"
      Appearance <- "CellSt1_25"
   Rectangle "cel_27" at 216,290 size 78x45
      Appearance <- "CellSt1_26"
   IOField "io_29" at 221,296 size 68x33; FormatPattern 999
      ProcessValue <- "Cell1_26"
      Appearance <- "CellSt1_26"
   Rectangle "cel_28" at 216,340 size 78x45
      Appearance <- "CellSt1_27"
   IOField "io_30" at 221,346 size 68x33; FormatPattern 999
      ProcessValue <- "Cell1_27"
      Appearance <- "CellSt1_27"
   Rectangle "cel_29" at 216,390 size 78x45
      Appearance <- "CellSt1_28"
   IOField "io_31" at 221,396 size 68x33; FormatPattern 999
      ProcessValue <- "Cell1_28"
      Appearance <- "CellSt1_28"
   Rectangle "cel_30" at 216,440 size 78x45
      Appearance <- "CellSt1_29"
   IOField "io_32" at 221,446 size 68x33; FormatPattern 999
      ProcessValue <- "Cell1_29"
      Appearance <- "CellSt1_29"
   Rectangle "cel_31" at 216,490 size 78x45
      Appearance <- "CellSt1_30"
   IOField "io_33" at 221,496 size 68x33; FormatPattern 999
      ProcessValue <- "Cell1_30"
      Appearance <- "CellSt1_30"
   Rectangle "cel_32" at 216,540 size 78x45
      Appearance <- "CellSt1_31"
   IOField "io_34" at 221,546 size 68x33; FormatPattern 999
      ProcessValue <- "Cell1_31"
      Appearance <- "CellSt1_31"
   Rectangle "cel_33" at 216,590 size 78x45
      Appearance <- "CellSt1_32"
   IOField "io_35" at 221,596 size 68x33; FormatPattern 999
      ProcessValue <- "Cell1_32"
      Appearance <- "CellSt1_32"
   Rectangle "cel_34" at 216,640 size 78x45
      Appearance <- "CellSt1_33"
   IOField "io_36" at 221,646 size 68x33; FormatPattern 999
      ProcessValue <- "Cell1_33"
      Appearance <- "CellSt1_33"
   Rectangle "cel_35" at 216,690 size 78x45
      Appearance <- "CellSt1_34"
   IOField "io_37" at 221,696 size 68x33; FormatPattern 999
      ProcessValue <- "Cell1_34"
      Appearance <- "CellSt1_34"
   Rectangle "cel_36" at 216,740 size 78x45
      Appearance <- "CellSt1_35"
   IOField "io_38" at 221,746 size 68x33; FormatPattern 999
      ProcessValue <- "Cell1_35"
      Appearance <- "CellSt1_35"
   Rectangle "cel_37" at 302,190 size 78x45
      Appearance <- "CellSt1_36"
   IOField "io_39" at 307,196 size 68x33; FormatPattern 999
      ProcessValue <- "Cell1_36"
      Appearance <- "CellSt1_36"
   Rectangle "cel_38" at 302,240 size 78x45
      Appearance <- "CellSt1_37"
   IOField "io_40" at 307,246 size 68x33; FormatPattern 999
      ProcessValue <- "Cell1_37"
      Appearance <- "CellSt1_37"
   Rectangle "cel_39" at 302,290 size 78x45
      Appearance <- "CellSt1_38"
   IOField "io_41" at 307,296 size 68x33; FormatPattern 999
      ProcessValue <- "Cell1_38"
      Appearance <- "CellSt1_38"
   Rectangle "cel_40" at 302,340 size 78x45
      Appearance <- "CellSt1_39"
   IOField "io_42" at 307,346 size 68x33; FormatPattern 999
      ProcessValue <- "Cell1_39"
      Appearance <- "CellSt1_39"
   Rectangle "cel_41" at 302,390 size 78x45
      Appearance <- "CellSt1_40"
   IOField "io_43" at 307,396 size 68x33; FormatPattern 999
      ProcessValue <- "Cell1_40"
      Appearance <- "CellSt1_40"
   Rectangle "cel_42" at 302,440 size 78x45
      Appearance <- "CellSt1_41"
   IOField "io_44" at 307,446 size 68x33; FormatPattern 999
      ProcessValue <- "Cell1_41"
      Appearance <- "CellSt1_41"
   Rectangle "cel_43" at 302,490 size 78x45
      Appearance <- "CellSt1_42"
   IOField "io_45" at 307,496 size 68x33; FormatPattern 999
      ProcessValue <- "Cell1_42"
      Appearance <- "CellSt1_42"
   Rectangle "cel_44" at 302,540 size 78x45
      Appearance <- "CellSt1_43"
   IOField "io_46" at 307,546 size 68x33; FormatPattern 999
      ProcessValue <- "Cell1_43"
      Appearance <- "CellSt1_43"
   Rectangle "cel_45" at 302,590 size 78x45
      Appearance <- "CellSt1_44"
   IOField "io_47" at 307,596 size 68x33; FormatPattern 999
      ProcessValue <- "Cell1_44"
      Appearance <- "CellSt1_44"
   Rectangle "cel_46" at 302,640 size 78x45
      Appearance <- "CellSt1_45"
   IOField "io_48" at 307,646 size 68x33; FormatPattern 999
      ProcessValue <- "Cell1_45"
      Appearance <- "CellSt1_45"
   Rectangle "cel_47" at 302,690 size 78x45
      Appearance <- "CellSt1_46"
   IOField "io_49" at 307,696 size 68x33; FormatPattern 999
      ProcessValue <- "Cell1_46"
      Appearance <- "CellSt1_46"
   Rectangle "cel_48" at 302,740 size 78x45
      Appearance <- "CellSt1_47"
   IOField "io_50" at 307,746 size 68x33; FormatPattern 999
      ProcessValue <- "Cell1_47"
      Appearance <- "CellSt1_47"
   Rectangle "cel_49" at 558,190 size 78x45
      Appearance <- "CellSt0_00"
   IOField "io_51" at 563,196 size 68x33; FormatPattern 999
      ProcessValue <- "Cell0_00"
      Appearance <- "CellSt0_00"
   Rectangle "cel_50" at 558,240 size 78x45
      Appearance <- "CellSt0_01"
   IOField "io_52" at 563,246 size 68x33; FormatPattern 999
      ProcessValue <- "Cell0_01"
      Appearance <- "CellSt0_01"
   Rectangle "cel_51" at 558,290 size 78x45
      Appearance <- "CellSt0_02"
   IOField "io_53" at 563,296 size 68x33; FormatPattern 999
      ProcessValue <- "Cell0_02"
      Appearance <- "CellSt0_02"
   Rectangle "cel_52" at 558,340 size 78x45
      Appearance <- "CellSt0_03"
   IOField "io_54" at 563,346 size 68x33; FormatPattern 999
      ProcessValue <- "Cell0_03"
      Appearance <- "CellSt0_03"
   Rectangle "cel_53" at 558,390 size 78x45
      Appearance <- "CellSt0_04"
   IOField "io_55" at 563,396 size 68x33; FormatPattern 999
      ProcessValue <- "Cell0_04"
      Appearance <- "CellSt0_04"
   Rectangle "cel_54" at 558,440 size 78x45
      Appearance <- "CellSt0_05"
   IOField "io_56" at 563,446 size 68x33; FormatPattern 999
      ProcessValue <- "Cell0_05"
      Appearance <- "CellSt0_05"
   Rectangle "cel_55" at 558,490 size 78x45
      Appearance <- "CellSt0_06"
   IOField "io_57" at 563,496 size 68x33; FormatPattern 999
      ProcessValue <- "Cell0_06"
      Appearance <- "CellSt0_06"
   Rectangle "cel_56" at 558,540 size 78x45
      Appearance <- "CellSt0_07"
   IOField "io_58" at 563,546 size 68x33; FormatPattern 999
      ProcessValue <- "Cell0_07"
      Appearance <- "CellSt0_07"
   Rectangle "cel_57" at 558,590 size 78x45
      Appearance <- "CellSt0_08"
   IOField "io_59" at 563,596 size 68x33; FormatPattern 999
      ProcessValue <- "Cell0_08"
      Appearance <- "CellSt0_08"
   Rectangle "cel_58" at 558,640 size 78x45
      Appearance <- "CellSt0_09"
   IOField "io_60" at 563,646 size 68x33; FormatPattern 999
      ProcessValue <- "Cell0_09"
      Appearance <- "CellSt0_09"
   Rectangle "cel_59" at 558,690 size 78x45
      Appearance <- "CellSt0_10"
   IOField "io_61" at 563,696 size 68x33; FormatPattern 999
      ProcessValue <- "Cell0_10"
      Appearance <- "CellSt0_10"
   Rectangle "cel_60" at 558,740 size 78x45
      Appearance <- "CellSt0_11"
   IOField "io_62" at 563,746 size 68x33; FormatPattern 999
      ProcessValue <- "Cell0_11"
      Appearance <- "CellSt0_11"
   Rectangle "cel_61" at 644,190 size 78x45
      Appearance <- "CellSt0_12"
   IOField "io_63" at 649,196 size 68x33; FormatPattern 999
      ProcessValue <- "Cell0_12"
      Appearance <- "CellSt0_12"
   Rectangle "cel_62" at 644,240 size 78x45
      Appearance <- "CellSt0_13"
   IOField "io_64" at 649,246 size 68x33; FormatPattern 999
      ProcessValue <- "Cell0_13"
      Appearance <- "CellSt0_13"
   Rectangle "cel_63" at 644,290 size 78x45
      Appearance <- "CellSt0_14"
   IOField "io_65" at 649,296 size 68x33; FormatPattern 999
      ProcessValue <- "Cell0_14"
      Appearance <- "CellSt0_14"
   Rectangle "cel_64" at 644,340 size 78x45
      Appearance <- "CellSt0_15"
   IOField "io_66" at 649,346 size 68x33; FormatPattern 999
      ProcessValue <- "Cell0_15"
      Appearance <- "CellSt0_15"
   Rectangle "cel_65" at 644,390 size 78x45
      Appearance <- "CellSt0_16"
   IOField "io_67" at 649,396 size 68x33; FormatPattern 999
      ProcessValue <- "Cell0_16"
      Appearance <- "CellSt0_16"
   Rectangle "cel_66" at 644,440 size 78x45
      Appearance <- "CellSt0_17"
   IOField "io_68" at 649,446 size 68x33; FormatPattern 999
      ProcessValue <- "Cell0_17"
      Appearance <- "CellSt0_17"
   Rectangle "cel_67" at 644,490 size 78x45
      Appearance <- "CellSt0_18"
   IOField "io_69" at 649,496 size 68x33; FormatPattern 999
      ProcessValue <- "Cell0_18"
      Appearance <- "CellSt0_18"
   Rectangle "cel_68" at 644,540 size 78x45
      Appearance <- "CellSt0_19"
   IOField "io_70" at 649,546 size 68x33; FormatPattern 999
      ProcessValue <- "Cell0_19"
      Appearance <- "CellSt0_19"
   Rectangle "cel_69" at 644,590 size 78x45
      Appearance <- "CellSt0_20"
   IOField "io_71" at 649,596 size 68x33; FormatPattern 999
      ProcessValue <- "Cell0_20"
      Appearance <- "CellSt0_20"
   Rectangle "cel_70" at 644,640 size 78x45
      Appearance <- "CellSt0_21"
   IOField "io_72" at 649,646 size 68x33; FormatPattern 999
      ProcessValue <- "Cell0_21"
      Appearance <- "CellSt0_21"
   Rectangle "cel_71" at 644,690 size 78x45
      Appearance <- "CellSt0_22"
   IOField "io_73" at 649,696 size 68x33; FormatPattern 999
      ProcessValue <- "Cell0_22"
      Appearance <- "CellSt0_22"
   Rectangle "cel_72" at 644,740 size 78x45
      Appearance <- "CellSt0_23"
   IOField "io_74" at 649,746 size 68x33; FormatPattern 999
      ProcessValue <- "Cell0_23"
      Appearance <- "CellSt0_23"
   Rectangle "cel_73" at 729,190 size 78x45
      Appearance <- "CellSt0_24"
   IOField "io_75" at 734,196 size 68x33; FormatPattern 999
      ProcessValue <- "Cell0_24"
      Appearance <- "CellSt0_24"
   Rectangle "cel_74" at 729,240 size 78x45
      Appearance <- "CellSt0_25"
   IOField "io_76" at 734,246 size 68x33; FormatPattern 999
      ProcessValue <- "Cell0_25"
      Appearance <- "CellSt0_25"
   Rectangle "cel_75" at 729,290 size 78x45
      Appearance <- "CellSt0_26"
   IOField "io_77" at 734,296 size 68x33; FormatPattern 999
      ProcessValue <- "Cell0_26"
      Appearance <- "CellSt0_26"
   Rectangle "cel_76" at 729,340 size 78x45
      Appearance <- "CellSt0_27"
   IOField "io_78" at 734,346 size 68x33; FormatPattern 999
      ProcessValue <- "Cell0_27"
      Appearance <- "CellSt0_27"
   Rectangle "cel_77" at 729,390 size 78x45
      Appearance <- "CellSt0_28"
   IOField "io_79" at 734,396 size 68x33; FormatPattern 999
      ProcessValue <- "Cell0_28"
      Appearance <- "CellSt0_28"
   Rectangle "cel_78" at 729,440 size 78x45
      Appearance <- "CellSt0_29"
   IOField "io_80" at 734,446 size 68x33; FormatPattern 999
      ProcessValue <- "Cell0_29"
      Appearance <- "CellSt0_29"
   Rectangle "cel_79" at 729,490 size 78x45
      Appearance <- "CellSt0_30"
   IOField "io_81" at 734,496 size 68x33; FormatPattern 999
      ProcessValue <- "Cell0_30"
      Appearance <- "CellSt0_30"
   Rectangle "cel_80" at 729,540 size 78x45
      Appearance <- "CellSt0_31"
   IOField "io_82" at 734,546 size 68x33; FormatPattern 999
      ProcessValue <- "Cell0_31"
      Appearance <- "CellSt0_31"
   Rectangle "cel_81" at 729,590 size 78x45
      Appearance <- "CellSt0_32"
   IOField "io_83" at 734,596 size 68x33; FormatPattern 999
      ProcessValue <- "Cell0_32"
      Appearance <- "CellSt0_32"
   Rectangle "cel_82" at 729,640 size 78x45
      Appearance <- "CellSt0_33"
   IOField "io_84" at 734,646 size 68x33; FormatPattern 999
      ProcessValue <- "Cell0_33"
      Appearance <- "CellSt0_33"
   Rectangle "cel_83" at 729,690 size 78x45
      Appearance <- "CellSt0_34"
   IOField "io_85" at 734,696 size 68x33; FormatPattern 999
      ProcessValue <- "Cell0_34"
      Appearance <- "CellSt0_34"
   Rectangle "cel_84" at 729,740 size 78x45
      Appearance <- "CellSt0_35"
   IOField "io_86" at 734,746 size 68x33; FormatPattern 999
      ProcessValue <- "Cell0_35"
      Appearance <- "CellSt0_35"
   Rectangle "cel_85" at 814,190 size 78x45
      Appearance <- "CellSt0_36"
   IOField "io_87" at 820,196 size 68x33; FormatPattern 999
      ProcessValue <- "Cell0_36"
      Appearance <- "CellSt0_36"
   Rectangle "cel_86" at 814,240 size 78x45
      Appearance <- "CellSt0_37"
   IOField "io_88" at 820,246 size 68x33; FormatPattern 999
      ProcessValue <- "Cell0_37"
      Appearance <- "CellSt0_37"
   Rectangle "cel_87" at 814,290 size 78x45
      Appearance <- "CellSt0_38"
   IOField "io_89" at 820,296 size 68x33; FormatPattern 999
      ProcessValue <- "Cell0_38"
      Appearance <- "CellSt0_38"
   Rectangle "cel_88" at 814,340 size 78x45
      Appearance <- "CellSt0_39"
   IOField "io_90" at 820,346 size 68x33; FormatPattern 999
      ProcessValue <- "Cell0_39"
      Appearance <- "CellSt0_39"
   Rectangle "cel_89" at 814,390 size 78x45
      Appearance <- "CellSt0_40"
   IOField "io_91" at 820,396 size 68x33; FormatPattern 999
      ProcessValue <- "Cell0_40"
      Appearance <- "CellSt0_40"
   Rectangle "cel_90" at 814,440 size 78x45
      Appearance <- "CellSt0_41"
   IOField "io_92" at 820,446 size 68x33; FormatPattern 999
      ProcessValue <- "Cell0_41"
      Appearance <- "CellSt0_41"
   Rectangle "cel_91" at 814,490 size 78x45
      Appearance <- "CellSt0_42"
   IOField "io_93" at 820,496 size 68x33; FormatPattern 999
      ProcessValue <- "Cell0_42"
      Appearance <- "CellSt0_42"
   Rectangle "cel_92" at 814,540 size 78x45
      Appearance <- "CellSt0_43"
   IOField "io_94" at 820,546 size 68x33; FormatPattern 999
      ProcessValue <- "Cell0_43"
      Appearance <- "CellSt0_43"
   Rectangle "cel_93" at 814,590 size 78x45
      Appearance <- "CellSt0_44"
   IOField "io_95" at 820,596 size 68x33; FormatPattern 999
      ProcessValue <- "Cell0_44"
      Appearance <- "CellSt0_44"
   Rectangle "cel_94" at 814,640 size 78x45
      Appearance <- "CellSt0_45"
   IOField "io_96" at 820,646 size 68x33; FormatPattern 999
      ProcessValue <- "Cell0_45"
      Appearance <- "CellSt0_45"
   Rectangle "cel_95" at 814,690 size 78x45
      Appearance <- "CellSt0_46"
   IOField "io_97" at 820,696 size 68x33; FormatPattern 999
      ProcessValue <- "Cell0_46"
      Appearance <- "CellSt0_46"
   Rectangle "cel_96" at 814,740 size 78x45
      Appearance <- "CellSt0_47"
   IOField "io_98" at 820,746 size 68x33; FormatPattern 999
      ProcessValue <- "Cell0_47"
      Appearance <- "CellSt0_47"
   IOField "crn_1" at 46,157 size 75x27; FormatPattern 999
      ProcessValue <- "Carried"
      HorizontalMovement <- "CraneGX"
   Rectangle "crn_2" at 424,198 size 90x30
      VerticalMovement <- "CraneY"
   TextField "frm_6" at 915,128 size 513x250; Text 'Text'
   TextField "txt_26" at 924,133 size 480x23; Text 'RUČNA NAREDBA'
   TextField "txt_27" at 924,167 size 90x28; Text 'Naredba'
   SymbolicIOField "sym_1" at 1014,167 size 180x28; TextOff '0'; TextOn '1'; TextList "TL_Cmd"
      ProcessValue <- "ManCmd"
   TextField "txt_28" at 924,203 size 90x28; Text 'x (0-3)'
   IOField "io_99" at 1014,203 size 52x28; FormatPattern 9
      ProcessValue <- "ManX"
   TextField "txt_29" at 1080,203 size 68x28; Text 'y (0-11)'
   IOField "io_100" at 1148,203 size 52x28; FormatPattern 99
      ProcessValue <- "ManY"
   TextField "txt_30" at 924,240 size 90x28; Text 'Bay'
   SymbolicIOField "sym_2" at 1014,240 size 180x28; TextOff '0'; TextOn '1'; TextList "TL_Bay"
      ProcessValue <- "ManBay"
   Button "btn_1" at 1230,167 size 180x102; TextOff 'IZVRŠI'
      on Press: SetBit("BtnManExec")
   TextField "txt_31" at 924,275 size 495x18; Text 'PODIGNI/SPUSTI: lokacija dizalice. x/y/Bay: cilj pomaka.'
   TextField "txt_32" at 924,303 size 90x27; Text 'Dizalica x'
   IOField "io_101" at 1014,303 size 38x27; FormatPattern 9
      ProcessValue <- "CraneX"
   TextField "txt_33" at 1059,303 size 22x27; Text 'y'
   IOField "io_102" at 1082,303 size 38x27; FormatPattern 99
      ProcessValue <- "CraneY"
   TextField "txt_34" at 1185,303 size 52x27; Text 'Bay'
   SymbolicIOField "sym_3" at 1238,303 size 180x27; TextOff '0'; TextOn '1'; TextList "TL_Bay"
      ProcessValue <- "CraneBay"
   TextField "txt_35" at 924,337 size 90x27; Text 'Teret (ID)'
   IOField "io_103" at 1014,337 size 60x27; FormatPattern 999
      ProcessValue <- "Carried"
   Rectangle "lmp_1" at 1185,341 size 16x18
      Appearance <- "CraneBusy"
   TextField "txt_36" at 1204,337 size 82x27; Text 'zauzeta'
   TextField "frm_7" at 915,385 size 513x163; Text 'Text'
   TextField "txt_37" at 924,390 size 300x23; Text 'RAVNOTEŽA BRODA (Bay 0)'
   Rectangle "lmp_2" at 1238,393 size 16x18
      Appearance <- "BalOk"
   TextField "txt_38" at 1257,390 size 165x23; Text '|L - R| <= 5'
   TextField "txt_39" at 924,422 size 112x27; Text 'Lijevo x0-1'
   Bar "bar_1" at 1036,423 size 300x23; MinimumValue 0; MaximumValue 24
      ProcessValue <- "BalL"
   IOField "io_104" at 1342,422 size 45x27; FormatPattern 99
      ProcessValue <- "BalL"
   TextField "txt_40" at 924,455 size 112x27; Text 'Desno x2-3'
   Bar "bar_2" at 1036,457 size 300x23; MinimumValue 0; MaximumValue 24
      ProcessValue <- "BalR"
   IOField "io_105" at 1342,455 size 45x27; FormatPattern 99
      ProcessValue <- "BalR"
   TextField "txt_41" at 924,492 size 112x27; Text 'Razlika L-R'
   IOField "io_106" at 1036,492 size 52x27; FormatPattern s99
      ProcessValue <- "BalDiff"
   TextField "txt_42" at 1110,492 size 82x27; Text 'Pramac'
   IOField "io_107" at 1192,492 size 45x27; FormatPattern 99
      ProcessValue <- "BalF"
   TextField "txt_43" at 1260,492 size 75x27; Text 'Krma'
   IOField "io_108" at 1335,492 size 45x27; FormatPattern 99
      ProcessValue <- "BalA"
   TextField "frm_8" at 915,555 size 513x103; Text 'Text'
   TextField "txt_44" at 924,560 size 300x23; Text 'NAPREDAK'
   TextField "txt_45" at 924,588 size 68x27; Text 'Istovar'
   IOField "io_109" at 992,588 size 39x27; FormatPattern 99
      ProcessValue <- "UDone"
   IOField "io_110" at 1035,588 size 39x27; FormatPattern 99
      ProcessValue <- "UTotal"
   TextField "txt_46" at 1095,588 size 68x27; Text 'Ukrcaj'
   IOField "io_111" at 1162,588 size 39x27; FormatPattern 99
      ProcessValue <- "LDone"
   IOField "io_112" at 1206,588 size 39x27; FormatPattern 99
      ProcessValue <- "LTotal"
   TextField "txt_47" at 1268,588 size 30x27; Text 'N'
   IOField "io_113" at 1298,588 size 45x27; FormatPattern 99
      ProcessValue <- "N"
   TextField "txt_48" at 924,623 size 68x27; Text 'Plan #'
   IOField "io_114" at 992,623 size 30x27; FormatPattern 9
      ProcessValue <- "PlanVariant"
   Rectangle "lmp_3" at 1050,628 size 16x18
      Appearance <- "Initialized"
   TextField "txt_49" at 1070,623 size 112x27; Text 'inicijalizirano'
   Rectangle "lmp_4" at 1192,628 size 16x18
      Appearance <- "LampDone"
   TextField "txt_50" at 1212,623 size 112x27; Text 'završeno'
   TextField "frm_9" at 915,665 size 513x182; Text 'Text'
   TextField "txt_51" at 924,668 size 225x20; Text 'LEGENDA ĆELIJA'
   TextField "frm_10" at 924,693 size 34x23; Text 'Text'
   TextField "txt_52" at 964,693 size 210x23; Text '0 prazno'
   TextField "frm_11" at 924,730 size 34x23; Text 'Text'
   TextField "txt_53" at 964,730 size 210x23; Text '1 zauzeto'
   TextField "frm_12" at 924,767 size 34x23; Text 'Text'
   TextField "txt_54" at 964,767 size 210x23; Text '2 za istovar'
   TextField "frm_13" at 924,803 size 34x23; Text 'Text'
   TextField "txt_55" at 964,803 size 210x23; Text '3 za ukrcaj'
   TextField "frm_14" at 1176,693 size 34x23; Text 'Text'
   TextField "txt_56" at 1216,693 size 210x23; Text '4 prebačeno'
   TextField "frm_15" at 1176,730 size 34x23; Text 'Text'
   TextField "txt_57" at 1216,730 size 210x23; Text '5 trenutni izvor'
   TextField "frm_16" at 1176,767 size 34x23; Text 'Text'
   TextField "txt_58" at 1216,767 size 210x23; Text '6 trenutni cilj'
   TextField "frm_17" at 1176,803 size 34x23; Text 'Text'
   TextField "txt_59" at 1216,803 size 210x23; Text '7 neispravan ID'

screen "Score" 1440x900, template "Tpl"
   TextField "frm_1" at 12,128 size 675x350; Text 'Text'
   TextField "txt_1" at 21,133 size 645x23; Text 'FUNKCIJA CILJA J = 0.5*T/(N*76 s) + 0.5*M/(4N)'
   TextField "txt_2" at 248,163 size 128x25; Text 'M'
   TextField "txt_3" at 382,163 size 128x25; Text 'T [s]'
   TextField "txt_4" at 518,163 size 128x25; Text 'J'
   TextField "txt_5" at 21,195 size 225x28; Text 'M (pravilo zadatka), stvarno'
   IOField "io_1" at 248,195 size 112x28; FormatPattern 99999
      ProcessValue <- "M"
   IOField "io_2" at 382,195 size 112x28; FormatPattern 99999.9
      ProcessValue <- "T"
   IOField "io_3" at 518,195 size 112x28; FormatPattern 9.9999
      ProcessValue <- "J"
   TextField "txt_6" at 21,230 size 225x28; Text 'M (FB1 brojač, MD107)'
   IOField "io_4" at 248,230 size 112x28; FormatPattern 99999
      ProcessValue <- "MFb1"
   IOField "io_5" at 518,230 size 112x28; FormatPattern 9.9999
      ProcessValue <- "JFb1"
   TextField "txt_7" at 21,265 size 225x28; Text 'Planirani rezultat'
   IOField "io_6" at 248,265 size 112x28; FormatPattern 99999
      ProcessValue <- "PredM"
   IOField "io_7" at 382,265 size 112x28; FormatPattern 99999.9
      ProcessValue <- "PredT"
   IOField "io_8" at 518,265 size 112x28; FormatPattern 9.9999
      ProcessValue <- "PredJ"
   TextField "txt_8" at 21,310 size 645x23; Text 'OPTIMIZACIJA PLANA (FB11: pohlepni plan, zatim lokalno pretraživanje)'
   TextField "txt_9" at 21,340 size 225x28; Text 'J pohlepnog plana'
   IOField "io_9" at 246,340 size 112x28; FormatPattern 9.9999
      ProcessValue <- "PredJ0"
   TextField "txt_10" at 368,340 size 150x28; Text 'Poboljšanje [%]'
   IOField "io_10" at 518,340 size 112x28; FormatPattern 99.99
      ProcessValue <- "ImpGainPct"
   TextField "txt_11" at 21,375 size 225x28; Text 'J optimiziranog plana'
   IOField "io_11" at 246,375 size 112x28; FormatPattern 9.9999
      ProcessValue <- "PredJ"
   TextField "txt_12" at 368,375 size 150x28; Text 'Evaluacije'
   IOField "io_12" at 518,375 size 112x28; FormatPattern 99999
      ProcessValue <- "ImpEvals"
   TextField "txt_13" at 21,410 size 225x28; Text 'Donja granica J (dokazana)'
   IOField "io_13" at 246,410 size 112x28; FormatPattern 9.9999
      ProcessValue <- "LbJ"
   TextField "txt_14" at 368,410 size 150x28; Text 'Udaljenost [%]'
   IOField "io_14" at 518,410 size 112x28; FormatPattern 99.99
      ProcessValue <- "GapPct"
   TextField "txt_15" at 21,445 size 225x25; Text 'Napredak planiranja [%]'
   Bar "bar_1" at 248,447 size 270x22; MinimumValue 0; MaximumValue 100
      ProcessValue <- "PlanProgress"
   IOField "io_15" at 525,443 size 60x28; FormatPattern 999
      ProcessValue <- "PlanProgress"
   TextField "frm_2" at 699,128 size 729x350; Text 'Text'
   TextField "txt_16" at 708,133 size 705x23; Text 'POSTAVKE PLANERA'
   TextField "txt_17" at 708,167 size 195x28; Text 'Redoslijed (korišten)'
   SymbolicIOField "sym_1" at 903,167 size 285x28; TextOff '0'; TextOn '1'; TextList "TL_Order"
      ProcessValue <- "OrderModeAct"
   TextField "txt_18" at 708,202 size 195x28; Text 'Pobjednička varijanta'
   IOField "io_16" at 903,202 size 45x28; FormatPattern 9
      ProcessValue <- "PlanVariant"
   TextField "txt_19" at 708,237 size 195x28; Text 'N (liste)'
   IOField "io_17" at 903,237 size 60x28; FormatPattern 99
      ProcessValue <- "N"
   Rectangle "lmp_1" at 708,278 size 16x18
      Appearance <- "Planning"
   TextField "txt_20" at 729,272 size 225x28; Text 'planiranje u tijeku'
   TextField "txt_21" at 708,317 size 705x22; Text 'Donja granica: T >= 40 s po kontejneru + 6 s po stupcu minimalnog x-puta (zatvorena formula),'
   TextField "txt_22" at 708,338 size 705x22; Text 'M >= 4 po kontejneru. Nijedan plan ne može biti bolji od te vrijednosti.'
   TextField "txt_23" at 708,368 size 705x22; Text 'Lokalno pretraživanje: premještanje, zamjena i premještanje para transfera; fiksni broj evaluacija,'
   TextField "txt_24" at 708,390 size 705x22; Text 'deterministički, uz pravilo ravnoteže |L-R| <= 5 u svakom koraku. Plan nikad nije lošiji od pohlepnog.'

screen "Screen_1" 1440x900, template "Tpl"
   TextField "txt_1" at 45,128 size 334x23; Text 'BAY 1 - SKLADIŠTE (yard)'
   TextField "txt_2" at 558,128 size 334x23; Text 'BAY 0 - BROD (ship)'
   TextField "frm_1" at 42,155 size 854x30; Text 'Text'
   TextField "frm_2" at 417,187 size 105x602; Text 'Text'
   TextField "txt_3" at 417,792 size 105x18; Text 'OBALA / kran y'
   TextField "frm_3" at 39,183 size 346x608; Text 'Text'
   TextField "frm_4" at 552,183 size 346x608; Text 'Text'
   TextField "frm_5" at 724,183 size 3x608; Text 'Text'
   TextField "txt_4" at 12,203 size 30x18; Text 'y0'
   TextField "txt_5" at 12,253 size 30x18; Text 'y1'
   TextField "txt_6" at 12,303 size 30x18; Text 'y2'
   TextField "txt_7" at 12,353 size 30x18; Text 'y3'
   TextField "txt_8" at 12,403 size 30x18; Text 'y4'
   TextField "txt_9" at 12,453 size 30x18; Text 'y5'
   TextField "txt_10" at 12,503 size 30x18; Text 'y6'
   TextField "txt_11" at 12,553 size 30x18; Text 'y7'
   TextField "txt_12" at 12,603 size 30x18; Text 'y8'
   TextField "txt_13" at 12,653 size 30x18; Text 'y9'
   TextField "txt_14" at 12,703 size 30x18; Text 'y10'
   TextField "txt_15" at 12,753 size 30x18; Text 'y11'
   TextField "txt_16" at 45,793 size 78x17; Text 'x0'
   TextField "txt_17" at 130,793 size 78x17; Text 'x1'
   TextField "txt_18" at 216,793 size 78x17; Text 'x2'
   TextField "txt_19" at 302,793 size 78x17; Text 'x3'
   TextField "txt_20" at 558,793 size 78x17; Text 'x0'
   TextField "txt_21" at 644,793 size 78x17; Text 'x1'
   TextField "txt_22" at 729,793 size 78x17; Text 'x2'
   TextField "txt_23" at 814,793 size 78x17; Text 'x3'
   TextField "txt_24" at 558,813 size 90x23; Text 'LIJEVO'
   IOField "io_1" at 648,813 size 45x23; FormatPattern 99
      ProcessValue <- "BalL"
   TextField "txt_25" at 729,813 size 90x23; Text 'DESNO'
   IOField "io_2" at 819,813 size 45x23; FormatPattern 99
      ProcessValue <- "BalR"
   Rectangle "cel_1" at 45,190 size 78x45
      Appearance <- "CellSt1_00"
   IOField "io_3" at 50,196 size 68x33; FormatPattern 999
      ProcessValue <- "Cell1_00"
      Appearance <- "CellSt1_00"
   Rectangle "cel_2" at 45,240 size 78x45
      Appearance <- "CellSt1_01"
   IOField "io_4" at 50,246 size 68x33; FormatPattern 999
      ProcessValue <- "Cell1_01"
      Appearance <- "CellSt1_01"
   Rectangle "cel_3" at 45,290 size 78x45
      Appearance <- "CellSt1_02"
   IOField "io_5" at 50,296 size 68x33; FormatPattern 999
      ProcessValue <- "Cell1_02"
      Appearance <- "CellSt1_02"
   Rectangle "cel_4" at 45,340 size 78x45
      Appearance <- "CellSt1_03"
   IOField "io_6" at 50,346 size 68x33; FormatPattern 999
      ProcessValue <- "Cell1_03"
      Appearance <- "CellSt1_03"
   Rectangle "cel_5" at 45,390 size 78x45
      Appearance <- "CellSt1_04"
   IOField "io_7" at 50,396 size 68x33; FormatPattern 999
      ProcessValue <- "Cell1_04"
      Appearance <- "CellSt1_04"
   Rectangle "cel_6" at 45,440 size 78x45
      Appearance <- "CellSt1_05"
   IOField "io_8" at 50,446 size 68x33; FormatPattern 999
      ProcessValue <- "Cell1_05"
      Appearance <- "CellSt1_05"
   Rectangle "cel_7" at 45,490 size 78x45
      Appearance <- "CellSt1_06"
   IOField "io_9" at 50,496 size 68x33; FormatPattern 999
      ProcessValue <- "Cell1_06"
      Appearance <- "CellSt1_06"
   Rectangle "cel_8" at 45,540 size 78x45
      Appearance <- "CellSt1_07"
   IOField "io_10" at 50,546 size 68x33; FormatPattern 999
      ProcessValue <- "Cell1_07"
      Appearance <- "CellSt1_07"
   Rectangle "cel_9" at 45,590 size 78x45
      Appearance <- "CellSt1_08"
   IOField "io_11" at 50,596 size 68x33; FormatPattern 999
      ProcessValue <- "Cell1_08"
      Appearance <- "CellSt1_08"
   Rectangle "cel_10" at 45,640 size 78x45
      Appearance <- "CellSt1_09"
   IOField "io_12" at 50,646 size 68x33; FormatPattern 999
      ProcessValue <- "Cell1_09"
      Appearance <- "CellSt1_09"
   Rectangle "cel_11" at 45,690 size 78x45
      Appearance <- "CellSt1_10"
   IOField "io_13" at 50,696 size 68x33; FormatPattern 999
      ProcessValue <- "Cell1_10"
      Appearance <- "CellSt1_10"
   Rectangle "cel_12" at 45,740 size 78x45
      Appearance <- "CellSt1_11"
   IOField "io_14" at 50,746 size 68x33; FormatPattern 999
      ProcessValue <- "Cell1_11"
      Appearance <- "CellSt1_11"
   Rectangle "cel_13" at 130,190 size 78x45
      Appearance <- "CellSt1_12"
   IOField "io_15" at 136,196 size 68x33; FormatPattern 999
      ProcessValue <- "Cell1_12"
      Appearance <- "CellSt1_12"
   Rectangle "cel_14" at 130,240 size 78x45
      Appearance <- "CellSt1_13"
   IOField "io_16" at 136,246 size 68x33; FormatPattern 999
      ProcessValue <- "Cell1_13"
      Appearance <- "CellSt1_13"
   Rectangle "cel_15" at 130,290 size 78x45
      Appearance <- "CellSt1_14"
   IOField "io_17" at 136,296 size 68x33; FormatPattern 999
      ProcessValue <- "Cell1_14"
      Appearance <- "CellSt1_14"
   Rectangle "cel_16" at 130,340 size 78x45
      Appearance <- "CellSt1_15"
   IOField "io_18" at 136,346 size 68x33; FormatPattern 999
      ProcessValue <- "Cell1_15"
      Appearance <- "CellSt1_15"
   Rectangle "cel_17" at 130,390 size 78x45
      Appearance <- "CellSt1_16"
   IOField "io_19" at 136,396 size 68x33; FormatPattern 999
      ProcessValue <- "Cell1_16"
      Appearance <- "CellSt1_16"
   Rectangle "cel_18" at 130,440 size 78x45
      Appearance <- "CellSt1_17"
   IOField "io_20" at 136,446 size 68x33; FormatPattern 999
      ProcessValue <- "Cell1_17"
      Appearance <- "CellSt1_17"
   Rectangle "cel_19" at 130,490 size 78x45
      Appearance <- "CellSt1_18"
   IOField "io_21" at 136,496 size 68x33; FormatPattern 999
      ProcessValue <- "Cell1_18"
      Appearance <- "CellSt1_18"
   Rectangle "cel_20" at 130,540 size 78x45
      Appearance <- "CellSt1_19"
   IOField "io_22" at 136,546 size 68x33; FormatPattern 999
      ProcessValue <- "Cell1_19"
      Appearance <- "CellSt1_19"
   Rectangle "cel_21" at 130,590 size 78x45
      Appearance <- "CellSt1_20"
   IOField "io_23" at 136,596 size 68x33; FormatPattern 999
      ProcessValue <- "Cell1_20"
      Appearance <- "CellSt1_20"
   Rectangle "cel_22" at 130,640 size 78x45
      Appearance <- "CellSt1_21"
   IOField "io_24" at 136,646 size 68x33; FormatPattern 999
      ProcessValue <- "Cell1_21"
      Appearance <- "CellSt1_21"
   Rectangle "cel_23" at 130,690 size 78x45
      Appearance <- "CellSt1_22"
   IOField "io_25" at 136,696 size 68x33; FormatPattern 999
      ProcessValue <- "Cell1_22"
      Appearance <- "CellSt1_22"
   Rectangle "cel_24" at 130,740 size 78x45
      Appearance <- "CellSt1_23"
   IOField "io_26" at 136,746 size 68x33; FormatPattern 999
      ProcessValue <- "Cell1_23"
      Appearance <- "CellSt1_23"
   Rectangle "cel_25" at 216,190 size 78x45
      Appearance <- "CellSt1_24"
   IOField "io_27" at 221,196 size 68x33; FormatPattern 999
      ProcessValue <- "Cell1_24"
      Appearance <- "CellSt1_24"
   Rectangle "cel_26" at 216,240 size 78x45
      Appearance <- "CellSt1_25"
   IOField "io_28" at 221,246 size 68x33; FormatPattern 999
      ProcessValue <- "Cell1_25"
      Appearance <- "CellSt1_25"
   Rectangle "cel_27" at 216,290 size 78x45
      Appearance <- "CellSt1_26"
   IOField "io_29" at 221,296 size 68x33; FormatPattern 999
      ProcessValue <- "Cell1_26"
      Appearance <- "CellSt1_26"
   Rectangle "cel_28" at 216,340 size 78x45
      Appearance <- "CellSt1_27"
   IOField "io_30" at 221,346 size 68x33; FormatPattern 999
      ProcessValue <- "Cell1_27"
      Appearance <- "CellSt1_27"
   Rectangle "cel_29" at 216,390 size 78x45
      Appearance <- "CellSt1_28"
   IOField "io_31" at 221,396 size 68x33; FormatPattern 999
      ProcessValue <- "Cell1_28"
      Appearance <- "CellSt1_28"
   Rectangle "cel_30" at 216,440 size 78x45
      Appearance <- "CellSt1_29"
   IOField "io_32" at 221,446 size 68x33; FormatPattern 999
      ProcessValue <- "Cell1_29"
      Appearance <- "CellSt1_29"
   Rectangle "cel_31" at 216,490 size 78x45
      Appearance <- "CellSt1_30"
   IOField "io_33" at 221,496 size 68x33; FormatPattern 999
      ProcessValue <- "Cell1_30"
      Appearance <- "CellSt1_30"
   Rectangle "cel_32" at 216,540 size 78x45
      Appearance <- "CellSt1_31"
   IOField "io_34" at 221,546 size 68x33; FormatPattern 999
      ProcessValue <- "Cell1_31"
      Appearance <- "CellSt1_31"
   Rectangle "cel_33" at 216,590 size 78x45
      Appearance <- "CellSt1_32"
   IOField "io_35" at 221,596 size 68x33; FormatPattern 999
      ProcessValue <- "Cell1_32"
      Appearance <- "CellSt1_32"
   Rectangle "cel_34" at 216,640 size 78x45
      Appearance <- "CellSt1_33"
   IOField "io_36" at 221,646 size 68x33; FormatPattern 999
      ProcessValue <- "Cell1_33"
      Appearance <- "CellSt1_33"
   Rectangle "cel_35" at 216,690 size 78x45
      Appearance <- "CellSt1_34"
   IOField "io_37" at 221,696 size 68x33; FormatPattern 999
      ProcessValue <- "Cell1_34"
      Appearance <- "CellSt1_34"
   Rectangle "cel_36" at 216,740 size 78x45
      Appearance <- "CellSt1_35"
   IOField "io_38" at 221,746 size 68x33; FormatPattern 999
      ProcessValue <- "Cell1_35"
      Appearance <- "CellSt1_35"
   Rectangle "cel_37" at 302,190 size 78x45
      Appearance <- "CellSt1_36"
   IOField "io_39" at 307,196 size 68x33; FormatPattern 999
      ProcessValue <- "Cell1_36"
      Appearance <- "CellSt1_36"
   Rectangle "cel_38" at 302,240 size 78x45
      Appearance <- "CellSt1_37"
   IOField "io_40" at 307,246 size 68x33; FormatPattern 999
      ProcessValue <- "Cell1_37"
      Appearance <- "CellSt1_37"
   Rectangle "cel_39" at 302,290 size 78x45
      Appearance <- "CellSt1_38"
   IOField "io_41" at 307,296 size 68x33; FormatPattern 999
      ProcessValue <- "Cell1_38"
      Appearance <- "CellSt1_38"
   Rectangle "cel_40" at 302,340 size 78x45
      Appearance <- "CellSt1_39"
   IOField "io_42" at 307,346 size 68x33; FormatPattern 999
      ProcessValue <- "Cell1_39"
      Appearance <- "CellSt1_39"
   Rectangle "cel_41" at 302,390 size 78x45
      Appearance <- "CellSt1_40"
   IOField "io_43" at 307,396 size 68x33; FormatPattern 999
      ProcessValue <- "Cell1_40"
      Appearance <- "CellSt1_40"
   Rectangle "cel_42" at 302,440 size 78x45
      Appearance <- "CellSt1_41"
   IOField "io_44" at 307,446 size 68x33; FormatPattern 999
      ProcessValue <- "Cell1_41"
      Appearance <- "CellSt1_41"
   Rectangle "cel_43" at 302,490 size 78x45
      Appearance <- "CellSt1_42"
   IOField "io_45" at 307,496 size 68x33; FormatPattern 999
      ProcessValue <- "Cell1_42"
      Appearance <- "CellSt1_42"
   Rectangle "cel_44" at 302,540 size 78x45
      Appearance <- "CellSt1_43"
   IOField "io_46" at 307,546 size 68x33; FormatPattern 999
      ProcessValue <- "Cell1_43"
      Appearance <- "CellSt1_43"
   Rectangle "cel_45" at 302,590 size 78x45
      Appearance <- "CellSt1_44"
   IOField "io_47" at 307,596 size 68x33; FormatPattern 999
      ProcessValue <- "Cell1_44"
      Appearance <- "CellSt1_44"
   Rectangle "cel_46" at 302,640 size 78x45
      Appearance <- "CellSt1_45"
   IOField "io_48" at 307,646 size 68x33; FormatPattern 999
      ProcessValue <- "Cell1_45"
      Appearance <- "CellSt1_45"
   Rectangle "cel_47" at 302,690 size 78x45
      Appearance <- "CellSt1_46"
   IOField "io_49" at 307,696 size 68x33; FormatPattern 999
      ProcessValue <- "Cell1_46"
      Appearance <- "CellSt1_46"
   Rectangle "cel_48" at 302,740 size 78x45
      Appearance <- "CellSt1_47"
   IOField "io_50" at 307,746 size 68x33; FormatPattern 999
      ProcessValue <- "Cell1_47"
      Appearance <- "CellSt1_47"
   Rectangle "cel_49" at 558,190 size 78x45
      Appearance <- "CellSt0_00"
   IOField "io_51" at 563,196 size 68x33; FormatPattern 999
      ProcessValue <- "Cell0_00"
      Appearance <- "CellSt0_00"
   Rectangle "cel_50" at 558,240 size 78x45
      Appearance <- "CellSt0_01"
   IOField "io_52" at 563,246 size 68x33; FormatPattern 999
      ProcessValue <- "Cell0_01"
      Appearance <- "CellSt0_01"
   Rectangle "cel_51" at 558,290 size 78x45
      Appearance <- "CellSt0_02"
   IOField "io_53" at 563,296 size 68x33; FormatPattern 999
      ProcessValue <- "Cell0_02"
      Appearance <- "CellSt0_02"
   Rectangle "cel_52" at 558,340 size 78x45
      Appearance <- "CellSt0_03"
   IOField "io_54" at 563,346 size 68x33; FormatPattern 999
      ProcessValue <- "Cell0_03"
      Appearance <- "CellSt0_03"
   Rectangle "cel_53" at 558,390 size 78x45
      Appearance <- "CellSt0_04"
   IOField "io_55" at 563,396 size 68x33; FormatPattern 999
      ProcessValue <- "Cell0_04"
      Appearance <- "CellSt0_04"
   Rectangle "cel_54" at 558,440 size 78x45
      Appearance <- "CellSt0_05"
   IOField "io_56" at 563,446 size 68x33; FormatPattern 999
      ProcessValue <- "Cell0_05"
      Appearance <- "CellSt0_05"
   Rectangle "cel_55" at 558,490 size 78x45
      Appearance <- "CellSt0_06"
   IOField "io_57" at 563,496 size 68x33; FormatPattern 999
      ProcessValue <- "Cell0_06"
      Appearance <- "CellSt0_06"
   Rectangle "cel_56" at 558,540 size 78x45
      Appearance <- "CellSt0_07"
   IOField "io_58" at 563,546 size 68x33; FormatPattern 999
      ProcessValue <- "Cell0_07"
      Appearance <- "CellSt0_07"
   Rectangle "cel_57" at 558,590 size 78x45
      Appearance <- "CellSt0_08"
   IOField "io_59" at 563,596 size 68x33; FormatPattern 999
      ProcessValue <- "Cell0_08"
      Appearance <- "CellSt0_08"
   Rectangle "cel_58" at 558,640 size 78x45
      Appearance <- "CellSt0_09"
   IOField "io_60" at 563,646 size 68x33; FormatPattern 999
      ProcessValue <- "Cell0_09"
      Appearance <- "CellSt0_09"
   Rectangle "cel_59" at 558,690 size 78x45
      Appearance <- "CellSt0_10"
   IOField "io_61" at 563,696 size 68x33; FormatPattern 999
      ProcessValue <- "Cell0_10"
      Appearance <- "CellSt0_10"
   Rectangle "cel_60" at 558,740 size 78x45
      Appearance <- "CellSt0_11"
   IOField "io_62" at 563,746 size 68x33; FormatPattern 999
      ProcessValue <- "Cell0_11"
      Appearance <- "CellSt0_11"
   Rectangle "cel_61" at 644,190 size 78x45
      Appearance <- "CellSt0_12"
   IOField "io_63" at 649,196 size 68x33; FormatPattern 999
      ProcessValue <- "Cell0_12"
      Appearance <- "CellSt0_12"
   Rectangle "cel_62" at 644,240 size 78x45
      Appearance <- "CellSt0_13"
   IOField "io_64" at 649,246 size 68x33; FormatPattern 999
      ProcessValue <- "Cell0_13"
      Appearance <- "CellSt0_13"
   Rectangle "cel_63" at 644,290 size 78x45
      Appearance <- "CellSt0_14"
   IOField "io_65" at 649,296 size 68x33; FormatPattern 999
      ProcessValue <- "Cell0_14"
      Appearance <- "CellSt0_14"
   Rectangle "cel_64" at 644,340 size 78x45
      Appearance <- "CellSt0_15"
   IOField "io_66" at 649,346 size 68x33; FormatPattern 999
      ProcessValue <- "Cell0_15"
      Appearance <- "CellSt0_15"
   Rectangle "cel_65" at 644,390 size 78x45
      Appearance <- "CellSt0_16"
   IOField "io_67" at 649,396 size 68x33; FormatPattern 999
      ProcessValue <- "Cell0_16"
      Appearance <- "CellSt0_16"
   Rectangle "cel_66" at 644,440 size 78x45
      Appearance <- "CellSt0_17"
   IOField "io_68" at 649,446 size 68x33; FormatPattern 999
      ProcessValue <- "Cell0_17"
      Appearance <- "CellSt0_17"
   Rectangle "cel_67" at 644,490 size 78x45
      Appearance <- "CellSt0_18"
   IOField "io_69" at 649,496 size 68x33; FormatPattern 999
      ProcessValue <- "Cell0_18"
      Appearance <- "CellSt0_18"
   Rectangle "cel_68" at 644,540 size 78x45
      Appearance <- "CellSt0_19"
   IOField "io_70" at 649,546 size 68x33; FormatPattern 999
      ProcessValue <- "Cell0_19"
      Appearance <- "CellSt0_19"
   Rectangle "cel_69" at 644,590 size 78x45
      Appearance <- "CellSt0_20"
   IOField "io_71" at 649,596 size 68x33; FormatPattern 999
      ProcessValue <- "Cell0_20"
      Appearance <- "CellSt0_20"
   Rectangle "cel_70" at 644,640 size 78x45
      Appearance <- "CellSt0_21"
   IOField "io_72" at 649,646 size 68x33; FormatPattern 999
      ProcessValue <- "Cell0_21"
      Appearance <- "CellSt0_21"
   Rectangle "cel_71" at 644,690 size 78x45
      Appearance <- "CellSt0_22"
   IOField "io_73" at 649,696 size 68x33; FormatPattern 999
      ProcessValue <- "Cell0_22"
      Appearance <- "CellSt0_22"
   Rectangle "cel_72" at 644,740 size 78x45
      Appearance <- "CellSt0_23"
   IOField "io_74" at 649,746 size 68x33; FormatPattern 999
      ProcessValue <- "Cell0_23"
      Appearance <- "CellSt0_23"
   Rectangle "cel_73" at 729,190 size 78x45
      Appearance <- "CellSt0_24"
   IOField "io_75" at 734,196 size 68x33; FormatPattern 999
      ProcessValue <- "Cell0_24"
      Appearance <- "CellSt0_24"
   Rectangle "cel_74" at 729,240 size 78x45
      Appearance <- "CellSt0_25"
   IOField "io_76" at 734,246 size 68x33; FormatPattern 999
      ProcessValue <- "Cell0_25"
      Appearance <- "CellSt0_25"
   Rectangle "cel_75" at 729,290 size 78x45
      Appearance <- "CellSt0_26"
   IOField "io_77" at 734,296 size 68x33; FormatPattern 999
      ProcessValue <- "Cell0_26"
      Appearance <- "CellSt0_26"
   Rectangle "cel_76" at 729,340 size 78x45
      Appearance <- "CellSt0_27"
   IOField "io_78" at 734,346 size 68x33; FormatPattern 999
      ProcessValue <- "Cell0_27"
      Appearance <- "CellSt0_27"
   Rectangle "cel_77" at 729,390 size 78x45
      Appearance <- "CellSt0_28"
   IOField "io_79" at 734,396 size 68x33; FormatPattern 999
      ProcessValue <- "Cell0_28"
      Appearance <- "CellSt0_28"
   Rectangle "cel_78" at 729,440 size 78x45
      Appearance <- "CellSt0_29"
   IOField "io_80" at 734,446 size 68x33; FormatPattern 999
      ProcessValue <- "Cell0_29"
      Appearance <- "CellSt0_29"
   Rectangle "cel_79" at 729,490 size 78x45
      Appearance <- "CellSt0_30"
   IOField "io_81" at 734,496 size 68x33; FormatPattern 999
      ProcessValue <- "Cell0_30"
      Appearance <- "CellSt0_30"
   Rectangle "cel_80" at 729,540 size 78x45
      Appearance <- "CellSt0_31"
   IOField "io_82" at 734,546 size 68x33; FormatPattern 999
      ProcessValue <- "Cell0_31"
      Appearance <- "CellSt0_31"
   Rectangle "cel_81" at 729,590 size 78x45
      Appearance <- "CellSt0_32"
   IOField "io_83" at 734,596 size 68x33; FormatPattern 999
      ProcessValue <- "Cell0_32"
      Appearance <- "CellSt0_32"
   Rectangle "cel_82" at 729,640 size 78x45
      Appearance <- "CellSt0_33"
   IOField "io_84" at 734,646 size 68x33; FormatPattern 999
      ProcessValue <- "Cell0_33"
      Appearance <- "CellSt0_33"
   Rectangle "cel_83" at 729,690 size 78x45
      Appearance <- "CellSt0_34"
   IOField "io_85" at 734,696 size 68x33; FormatPattern 999
      ProcessValue <- "Cell0_34"
      Appearance <- "CellSt0_34"
   Rectangle "cel_84" at 729,740 size 78x45
      Appearance <- "CellSt0_35"
   IOField "io_86" at 734,746 size 68x33; FormatPattern 999
      ProcessValue <- "Cell0_35"
      Appearance <- "CellSt0_35"
   Rectangle "cel_85" at 814,190 size 78x45
      Appearance <- "CellSt0_36"
   IOField "io_87" at 820,196 size 68x33; FormatPattern 999
      ProcessValue <- "Cell0_36"
      Appearance <- "CellSt0_36"
   Rectangle "cel_86" at 814,240 size 78x45
      Appearance <- "CellSt0_37"
   IOField "io_88" at 820,246 size 68x33; FormatPattern 999
      ProcessValue <- "Cell0_37"
      Appearance <- "CellSt0_37"
   Rectangle "cel_87" at 814,290 size 78x45
      Appearance <- "CellSt0_38"
   IOField "io_89" at 820,296 size 68x33; FormatPattern 999
      ProcessValue <- "Cell0_38"
      Appearance <- "CellSt0_38"
   Rectangle "cel_88" at 814,340 size 78x45
      Appearance <- "CellSt0_39"
   IOField "io_90" at 820,346 size 68x33; FormatPattern 999
      ProcessValue <- "Cell0_39"
      Appearance <- "CellSt0_39"
   Rectangle "cel_89" at 814,390 size 78x45
      Appearance <- "CellSt0_40"
   IOField "io_91" at 820,396 size 68x33; FormatPattern 999
      ProcessValue <- "Cell0_40"
      Appearance <- "CellSt0_40"
   Rectangle "cel_90" at 814,440 size 78x45
      Appearance <- "CellSt0_41"
   IOField "io_92" at 820,446 size 68x33; FormatPattern 999
      ProcessValue <- "Cell0_41"
      Appearance <- "CellSt0_41"
   Rectangle "cel_91" at 814,490 size 78x45
      Appearance <- "CellSt0_42"
   IOField "io_93" at 820,496 size 68x33; FormatPattern 999
      ProcessValue <- "Cell0_42"
      Appearance <- "CellSt0_42"
   Rectangle "cel_92" at 814,540 size 78x45
      Appearance <- "CellSt0_43"
   IOField "io_94" at 820,546 size 68x33; FormatPattern 999
      ProcessValue <- "Cell0_43"
      Appearance <- "CellSt0_43"
   Rectangle "cel_93" at 814,590 size 78x45
      Appearance <- "CellSt0_44"
   IOField "io_95" at 820,596 size 68x33; FormatPattern 999
      ProcessValue <- "Cell0_44"
      Appearance <- "CellSt0_44"
   Rectangle "cel_94" at 814,640 size 78x45
      Appearance <- "CellSt0_45"
   IOField "io_96" at 820,646 size 68x33; FormatPattern 999
      ProcessValue <- "Cell0_45"
      Appearance <- "CellSt0_45"
   Rectangle "cel_95" at 814,690 size 78x45
      Appearance <- "CellSt0_46"
   IOField "io_97" at 820,696 size 68x33; FormatPattern 999
      ProcessValue <- "Cell0_46"
      Appearance <- "CellSt0_46"
   Rectangle "cel_96" at 814,740 size 78x45
      Appearance <- "CellSt0_47"
   IOField "io_98" at 820,746 size 68x33; FormatPattern 999
      ProcessValue <- "Cell0_47"
      Appearance <- "CellSt0_47"
   IOField "crn_1" at 46,157 size 75x27; FormatPattern 999
      ProcessValue <- "Carried"
      HorizontalMovement <- "CraneGX"
   Rectangle "crn_2" at 424,198 size 90x30
      VerticalMovement <- "CraneY"
   TextField "frm_6" at 915,128 size 513x250; Text 'Text'
   TextField "txt_26" at 924,133 size 300x23; Text 'TRENUTNA NAREDBA'
   TextField "txt_27" at 924,163 size 90x27; Text 'Naredba'
   SymbolicIOField "sym_1" at 1014,163 size 165x27; TextOff '0'; TextOn '1'; TextList "TL_Cmd"
      ProcessValue <- "CurCmd"
   TextField "txt_28" at 1185,163 size 52x27; Text 'Vrsta'
   SymbolicIOField "sym_2" at 1238,163 size 180x27; TextOff '0'; TextOn '1'; TextList "TL_Kind"
      ProcessValue <- "CurKind"
   TextField "txt_29" at 924,197 size 90x27; Text 'Kontejner'
   IOField "io_99" at 1014,197 size 60x27; FormatPattern 999
      ProcessValue <- "CurId"
   TextField "txt_30" at 1185,197 size 52x27; Text 'Faza'
   SymbolicIOField "sym_3" at 1238,197 size 180x27; TextOff '0'; TextOn '1'; TextList "TL_Phase"
      ProcessValue <- "CurPhase"
   TextField "txt_31" at 924,230 size 90x27; Text 'Cilj x'
   IOField "io_100" at 1014,230 size 38x27; FormatPattern 9
      ProcessValue <- "CurX"
   TextField "txt_32" at 1059,230 size 22x27; Text 'y'
   IOField "io_101" at 1082,230 size 38x27; FormatPattern 99
      ProcessValue <- "CurY"
   TextField "txt_33" at 1185,230 size 52x27; Text 'Bay'
   SymbolicIOField "sym_4" at 1238,230 size 180x27; TextOff '0'; TextOn '1'; TextList "TL_Bay"
      ProcessValue <- "CurBay"
   TextField "txt_34" at 924,270 size 300x23; Text 'DIZALICA'
   TextField "txt_35" at 924,300 size 90x27; Text 'Položaj x'
   IOField "io_102" at 1014,300 size 38x27; FormatPattern 9
      ProcessValue <- "CraneX"
   TextField "txt_36" at 1059,300 size 22x27; Text 'y'
   IOField "io_103" at 1082,300 size 38x27; FormatPattern 99
      ProcessValue <- "CraneY"
   TextField "txt_37" at 1185,300 size 52x27; Text 'Bay'
   SymbolicIOField "sym_5" at 1238,300 size 180x27; TextOff '0'; TextOn '1'; TextList "TL_Bay"
      ProcessValue <- "CraneBay"
   TextField "txt_38" at 924,333 size 90x27; Text 'Teret (ID)'
   IOField "io_104" at 1014,333 size 60x27; FormatPattern 999
      ProcessValue <- "Carried"
   Rectangle "lmp_1" at 1185,338 size 16x18
      Appearance <- "CraneBusy"
   TextField "txt_39" at 1204,333 size 82x27; Text 'zauzeta'
   Rectangle "lmp_2" at 1290,338 size 16x18
      Appearance <- "Planning"
   TextField "txt_40" at 1310,333 size 112x27; Text 'planiranje'
   TextField "frm_7" at 915,385 size 513x163; Text 'Text'
   TextField "txt_41" at 924,390 size 300x23; Text 'RAVNOTEŽA BRODA (Bay 0)'
   Rectangle "lmp_3" at 1238,393 size 16x18
      Appearance <- "BalOk"
   TextField "txt_42" at 1257,390 size 165x23; Text '|L - R| <= 5'
   TextField "txt_43" at 924,422 size 112x27; Text 'Lijevo x0-1'
   Bar "bar_1" at 1036,423 size 300x23; MinimumValue 0; MaximumValue 24
      ProcessValue <- "BalL"
   IOField "io_105" at 1342,422 size 45x27; FormatPattern 99
      ProcessValue <- "BalL"
   TextField "txt_44" at 924,455 size 112x27; Text 'Desno x2-3'
   Bar "bar_2" at 1036,457 size 300x23; MinimumValue 0; MaximumValue 24
      ProcessValue <- "BalR"
   IOField "io_106" at 1342,455 size 45x27; FormatPattern 99
      ProcessValue <- "BalR"
   TextField "txt_45" at 924,492 size 112x27; Text 'Razlika L-R'
   IOField "io_107" at 1036,492 size 52x27; FormatPattern s99
      ProcessValue <- "BalDiff"
   TextField "txt_46" at 1110,492 size 82x27; Text 'Pramac'
   IOField "io_108" at 1192,492 size 45x27; FormatPattern 99
      ProcessValue <- "BalF"
   TextField "txt_47" at 1260,492 size 75x27; Text 'Krma'
   IOField "io_109" at 1335,492 size 45x27; FormatPattern 99
      ProcessValue <- "BalA"
   TextField "frm_8" at 915,555 size 513x103; Text 'Text'
   TextField "txt_48" at 924,560 size 300x23; Text 'NAPREDAK'
   TextField "txt_49" at 924,588 size 68x27; Text 'Istovar'
   IOField "io_110" at 992,588 size 39x27; FormatPattern 99
      ProcessValue <- "UDone"
   IOField "io_111" at 1035,588 size 39x27; FormatPattern 99
      ProcessValue <- "UTotal"
   TextField "txt_50" at 1095,588 size 68x27; Text 'Ukrcaj'
   IOField "io_112" at 1162,588 size 39x27; FormatPattern 99
      ProcessValue <- "LDone"
   IOField "io_113" at 1206,588 size 39x27; FormatPattern 99
      ProcessValue <- "LTotal"
   TextField "txt_51" at 1268,588 size 30x27; Text 'N'
   IOField "io_114" at 1298,588 size 45x27; FormatPattern 99
      ProcessValue <- "N"
   TextField "txt_52" at 924,623 size 68x27; Text 'Plan #'
   IOField "io_115" at 992,623 size 30x27; FormatPattern 9
      ProcessValue <- "PlanVariant"
   Rectangle "lmp_4" at 1050,628 size 16x18
      Appearance <- "Initialized"
   TextField "txt_53" at 1070,623 size 112x27; Text 'inicijalizirano'
   Rectangle "lmp_5" at 1192,628 size 16x18
      Appearance <- "LampDone"
   TextField "txt_54" at 1212,623 size 112x27; Text 'završeno'
   TextField "frm_9" at 915,665 size 513x182; Text 'Text'
   TextField "txt_55" at 924,668 size 225x20; Text 'LEGENDA ĆELIJA'
   TextField "frm_10" at 924,693 size 34x23; Text 'Text'
   TextField "txt_56" at 964,693 size 210x23; Text '0 prazno'
   TextField "frm_11" at 924,730 size 34x23; Text 'Text'
   TextField "txt_57" at 964,730 size 210x23; Text '1 zauzeto'
   TextField "frm_12" at 924,767 size 34x23; Text 'Text'
   TextField "txt_58" at 964,767 size 210x23; Text '2 za istovar'
   TextField "frm_13" at 924,803 size 34x23; Text 'Text'
   TextField "txt_59" at 964,803 size 210x23; Text '3 za ukrcaj'
   TextField "frm_14" at 1176,693 size 34x23; Text 'Text'
   TextField "txt_60" at 1216,693 size 210x23; Text '4 prebačeno'
   TextField "frm_15" at 1176,730 size 34x23; Text 'Text'
   TextField "txt_61" at 1216,730 size 210x23; Text '5 trenutni izvor'
   TextField "frm_16" at 1176,767 size 34x23; Text 'Text'
   TextField "txt_62" at 1216,767 size 210x23; Text '6 trenutni cilj'
   TextField "frm_17" at 1176,803 size 34x23; Text 'Text'
   TextField "txt_63" at 1216,803 size 210x23; Text '7 neispravan ID'
*)